(* Logix 5000 project; controller NWGG 1756-L72 rev 35.12; software revision 35.00; part 3 of 19 *)
(* tags used below, declared in another part *)
   _6Y : ALIAS FOR I25[2].3;
   _700_TREAT : ALIAS FOR I7.3;
   _709G_TREAT : ALIAS FOR B21[9].7;
   _9_DRIP_GAT : ALIAS FOR O24[7].7;
   _9_GATE_SV : ALIAS FOR O24[7].0;
   _9_GATE_SV1 : ALIAS FOR O24[7].1;
   _9_TREATER : ALIAS FOR I24[6].7;
   _9_TRT_MB : ALIAS FOR B3[9].0;
   _9_TRT_MOV : ALIAS FOR O24[7].4;
   _9_TRT_STB : ALIAS FOR B3[9].1;
   _9_TRT_STPB : ALIAS FOR B3[9].2;
   A16 : INT[250];
   A_ACC : ALIAS FOR N10[11];
   A_HOLD_B : ALIAS FOR B3[1].4;
   A_HOLD_MB : ALIAS FOR B3[1].3;
   A_HOLD_REL : ALIAS FOR B3[1].5;
   A_MAIN_CNT : ALIAS FOR C5[0].PRE;
   A_MAIN_CNT1 : ALIAS FOR C5[0].ACC;
   A_MAIN_TRE : ALIAS FOR C5[0];
   A_PRESET : ALIAS FOR N10[10];
   A_PRESET_S : ALIAS FOR N10[12];
   A_RESET_PB : ALIAS FOR B3[1].2;
   A_SET : ALIAS FOR B3[1].6;
   A_STB_AUTO : ALIAS FOR B3[1].0;
   A_STPB_AUT : ALIAS FOR B3[1].1;
   A_TREATER : ALIAS FOR I24[6].8;
   A_TREATER1 : ALIAS FOR T4[59];
   B15 : DINT[100];
   B17 : DINT[30];
   B21 : DINT[255];
   B3 : DINT[250];
   B9 : DINT[150];
   Beta : BOOL;
   C5 : COUNTER[50];
   F8 : REAL[27];
   I1 : ALIAS FOR R1S0_AENTR:1:I.Data;
   I1_000_Bit00 : ALIAS FOR I1.0;
   I1_000_Bit02 : ALIAS FOR I1.2;
   I1_000_Bit03 : ALIAS FOR I1.3;
   I1_000_Bit05 : ALIAS FOR I1.5;
   I1_000_Bit06 : ALIAS FOR I1.6;
   I1_000_Bit08 : ALIAS FOR I1.8;
   I1_000_Bit09 : ALIAS FOR I1.9;
   I1_000_Bit11 : ALIAS FOR I1.11;
   I1_000_Bit12 : ALIAS FOR I1.12;
   I1_000_Bit14 : ALIAS FOR I1.14;
   I2 : ALIAS FOR R1S0_AENTR:2:I.Data;
   I24_004_Bit00 : ALIAS FOR I24[4].0;
   I24_004_Bit01 : ALIAS FOR I24[4].1;
   I24_004_Bit02 : ALIAS FOR I24[4].2;
   I24_004_Bit03 : ALIAS FOR I24[4].3;
   I24_006_Bit13 : ALIAS FOR I24[6].13;
   I25_002_Bit04 : ALIAS FOR I25[2].4;
   I2_000_Bit00 : ALIAS FOR I2.0;
   I2_000_Bit02 : ALIAS FOR I2.2;
   I2_000_Bit03 : ALIAS FOR I2.3;
   I2_000_Bit05 : ALIAS FOR I2.5;
   I2_000_Bit06 : ALIAS FOR I2.6;
   I2_000_Bit08 : ALIAS FOR I2.8;
   I2_000_Bit09 : ALIAS FOR I2.9;
   I2_000_Bit11 : ALIAS FOR I2.11;
   I2_000_Bit12 : ALIAS FOR I2.12;
   I2_000_Bit14 : ALIAS FOR I2.14;
   I3 : ALIAS FOR R1S0_AENTR:3:I.Data;
   I3_000_Bit00 : ALIAS FOR I3.0;
   I3_000_Bit02 : ALIAS FOR I3.2;
   I3_000_Bit03 : ALIAS FOR I3.3;
   I3_000_Bit05 : ALIAS FOR I3.5;
   I3_000_Bit06 : ALIAS FOR I3.6;
   I3_000_Bit08 : ALIAS FOR I3.8;
   I3_000_Bit09 : ALIAS FOR I3.9;
   I3_000_Bit11 : ALIAS FOR I3.11;
   I3_000_Bit12 : ALIAS FOR I3.12;
   I3_000_Bit14 : ALIAS FOR I3.14;
   I4 : ALIAS FOR R1S0_AENTR:4:I.Data;
   I4_000_Bit00 : ALIAS FOR I4.0;
   I4_000_Bit02 : ALIAS FOR I4.2;
   I4_000_Bit04 : ALIAS FOR I4.4;
   InEUMax : REAL;
   MAIN_TIMER : ALIAS FOR T11[0];
   MAIN_TIMER1 : ALIAS FOR T11[1];
   N20 : DINT[30];
   N23 : DINT[5];
   N7 : DINT[100];
   O10 : ALIAS FOR R1S0_AENTR:10:O.Data;
   O11 : ALIAS FOR R1S0_AENTR:11:O.Data;
   O12 : ALIAS FOR R1S0_AENTR:12:O.Data;
   O24_005_Bit00 : ALIAS FOR O24[5].0;
   O24_005_Bit01 : ALIAS FOR O24[5].1;
   O24_005_Bit02 : ALIAS FOR O24[5].2;
   O24_007_Bit05 : ALIAS FOR O24[7].5;
   O25_010_Bit04 : ALIAS FOR O25[10].4;
   O25_010_Bit07 : ALIAS FOR O25[10].7;
   P1_AUTO_SE : ALIAS FOR B3[5].1;
   P1_RUN_AUT1 : ALIAS FOR B3[4].1;
   P1_SEC_SEL : ALIAS FOR B17[1].1;
   P2_AUTO_SE : ALIAS FOR B3[5].2;
   P2_RUN_AUT1 : ALIAS FOR B3[4].2;
   P2_SEC_SEL : ALIAS FOR B17[1].2;
   P3_AUTO_SE : ALIAS FOR B3[5].3;
   P3_RUN_AUT1 : ALIAS FOR B3[4].3;
   P3_SEC_SEL : ALIAS FOR B17[1].3;
   P4_AUTO_SE : ALIAS FOR B3[5].4;
   P4_RUN_AUT1 : ALIAS FOR B3[4].4;
   P4_SEC_SEL : ALIAS FOR B17[1].4;
   P_RESET_AU : ALIAS FOR B3[4].0;
   PUMP_NO_FL : ALIAS FOR B12[11].0;
   T11_AIRSG1 : ALIAS FOR T4[0];
   T11_AIRSG2 : ALIAS FOR T4[1];
   T11_AUTO_A : ALIAS FOR T4[61];
   T11_TREAT : ALIAS FOR B3[11].0;
   T11_TRT_MO : ALIAS FOR T4[41];
   T12_DLY_TR : ALIAS FOR T4[2];
   T12_DLY_TR3 : ALIAS FOR T4[3];
   T12_TREAT : ALIAS FOR B3[12].0;
   T12_TRT_MO : ALIAS FOR T4[42];
   T13_DLY_TR : ALIAS FOR T4[4];
   T13_DLY_TR3 : ALIAS FOR T4[5];
   T13_TREAT : ALIAS FOR B3[13].0;
   T13_TRT_MO : ALIAS FOR T4[43];
   T13C_TREAT : ALIAS FOR B21[70].10;
   T14_DLY_TR : ALIAS FOR T4[6];
   T14_DLY_TR3 : ALIAS FOR T4[7];
   T14_TREAT : ALIAS FOR B3[14].0;
   T14_TRT_MO : ALIAS FOR T4[44];
   T15_TREAT : ALIAS FOR B3[15].0;
   T15_TRT_MO : ALIAS FOR T4[45];
   T15_TRT_OF : ALIAS FOR T4[9];
   T15_TRT_ON : ALIAS FOR T4[8];
   T16_TREAT : ALIAS FOR B3[16].0;
   T16_TRT_MO : ALIAS FOR T4[46];
   T16_TRT_OF : ALIAS FOR T4[11];
   T16_TRT_ON : ALIAS FOR T4[10];

   T17_HOLD_A : ALIAS FOR B3[17].3;
   T17_HOLD_M : ALIAS FOR B3[17].6;
   T17_K_FACT : ALIAS FOR F8[13];
   T17_LOW_BI : ALIAS FOR B15[17].2;
   T17_METER : ALIAS FOR I2.5;
   T17_NO_PAS : ALIAS FOR B17[17].2;
   T17_NULL_V : ALIAS FOR A16[178];
   T17_NULL_V1 : ALIAS FOR A16[179];
   T17_OP_DEF : ALIAS FOR A16[176];
   T17_OP_DEF1 : ALIAS FOR A16[177];
   T17_OP_NAM : ALIAS FOR A16[173];
   T17_OP_NAM1 : ALIAS FOR A16[174];
   T17_OPEN_A : ALIAS FOR B3[17].8;
   T17_OPEN_M : ALIAS FOR O10.5;
   T17_OPEN_M1 : ALIAS FOR B3[17].10;
   T17_RELEAS : ALIAS FOR B3[17].5;
   T17_RESET : ALIAS FOR B3[17].7;
   T17_SET_AU : ALIAS FOR B3[17].2;
   T17_SET_DE : ALIAS FOR B3[2].6;
   T17_SET_LO : ALIAS FOR B3[17].13;
   T17_SET_MA : ALIAS FOR B3[17].12;
   T17_SET_NA : ALIAS FOR A16[170];
   T17_SET_NA1 : ALIAS FOR A16[171];
   T17_SET_NA2 : ALIAS FOR B17[17].0;
   T17_STOP_A : ALIAS FOR B3[17].4;
   T17_TREAT : ALIAS FOR B3[17].0;
   T17_TRT_MO : ALIAS FOR T4[47];
   T17_TRT_MO1 : ALIAS FOR T4[47].PRE;
   T17_TRT_MO2 : ALIAS FOR T4[47].ACC;
   T17_TRT_OF : ALIAS FOR T4[13];
   T17_TRT_OF1 : ALIAS FOR T4[13].PRE;
   T17_TRT_OF2 : ALIAS FOR T4[13].ACC;
   T17_TRT_ON : ALIAS FOR T4[12];
   T17_TRT_ON1 : ALIAS FOR T4[12].PRE;
   T17_TRT_ON2 : ALIAS FOR T4[12].ACC;
   T19 : TIMER[2] := ([0].PRE := 11000, [0].ACC := 11000, [1].PRE := 60000, [1].ACC := 60000);
   T19C_AIR_G : ALIAS FOR O12.13;
   T19C_AIR_S : ALIAS FOR B21[71].11;
   T19C_CLOSE : ALIAS FOR O12.12;
   T19C_CLOSE1 : ALIAS FOR T22[3];
   T19C_CLOSE2 : ALIAS FOR T22[3].PRE;
   T19C_CLOSE3 : ALIAS FOR T22[3].ACC;
   T19C_GATE : ALIAS FOR B21[71].0;
   T19C_GATE1 : ALIAS FOR B21[71].1;
   T19C_GATE2 : ALIAS FOR B21[71].3;
   T19C_GATE3 : ALIAS FOR B21[71].4;
   T19C_GATE4 : ALIAS FOR B21[71].5;
   T19C_GATE5 : ALIAS FOR B21[71].6;
   T19C_GATE6 : ALIAS FOR B21[71].7;
   T19C_GATE7 : ALIAS FOR B21[71].8;
   T19C_GATE8 : ALIAS FOR B21[71].9;
   T19C_GATEC : ALIAS FOR B21[71].2;
   T19C_GATET : ALIAS FOR C5[4];
   T19C_OPEN : ALIAS FOR O12.11;
   T19C_SET_D : ALIAS FOR B21[71].14;
   T19C_TMR_A : ALIAS FOR C5[4].ACC;
   T19C_TMR_P : ALIAS FOR C5[4].PRE;
   T19C_TREAT : ALIAS FOR B21[71].10;
   T19C_TRT_M : ALIAS FOR T22[4];
   T19C_TRT_M1 : ALIAS FOR T22[4].PRE;
   T19C_TRT_M2 : ALIAS FOR T22[4].ACC;
   T19C_TRT_O : ALIAS FOR T22[0];
   T19C_TRT_O1 : ALIAS FOR T22[0].PRE;
   T19C_TRT_O2 : ALIAS FOR T22[0].ACC;
   T21_AIR_GA : ALIAS FOR I2.6;
   T21_AIR_SV : ALIAS FOR O10.6;
   T21_ASCII : ALIAS FOR B17[21].1;
   T21_ASSII : ALIAS FOR A16[212];
   T21_ASSII1 : ALIAS FOR A16[215];
   T21_AUTO_A : ALIAS FOR T4[71];
   T21_AUTO_A1 : ALIAS FOR T4[71].PRE;
   T21_AUTO_A2 : ALIAS FOR T4[71].ACC;
   T21_AUTO_M : ALIAS FOR B3[21].1;
   T21_AUTO_S : ALIAS FOR B3[21].14;
   T21_BINDIC : ALIAS FOR I1.1;
   T21_CAL_CL : ALIAS FOR B15[61].3;
   T21_CAL_LA : ALIAS FOR B15[61].2;
   T21_CAL_OP : ALIAS FOR B15[61].4;
   T21_CAL_ST : ALIAS FOR B15[61].1;
   T21_CLOSE : ALIAS FOR O10.7;
   T21_CLOSE1 : ALIAS FOR B3[21].9;
   T21_CLOSE2 : ALIAS FOR B3[21].11;
   T21_CORREC : ALIAS FOR F8[16];
   T21_FAULT : ALIAS FOR B3[21].15;
   T21_GATE_C : ALIAS FOR C5[21];
   T21_GATE_C1 : ALIAS FOR C5[21].PRE;
   T21_GATE_C2 : ALIAS FOR C5[21].ACC;
   T21_HOLD_A : ALIAS FOR B3[21].3;
   T21_HOLD_M : ALIAS FOR B3[21].6;
   T21_K_FACT : ALIAS FOR F8[15];
   T21_LOW_BI : ALIAS FOR B15[21].2;
   T21_METER : ALIAS FOR I2.8;
   T21_MOVE_D : ALIAS FOR I2.7;
   T21_NO_PAS : ALIAS FOR B17[21].2;
   T21_NULL_V : ALIAS FOR A16[218];
   T21_NULL_V1 : ALIAS FOR A16[219];
   T21_OP_DEF : ALIAS FOR A16[216];
   T21_OP_DEF1 : ALIAS FOR A16[217];
   T21_OP_NAM : ALIAS FOR A16[213];
   T21_OP_NAM1 : ALIAS FOR A16[214];
   T21_OPEN_A : ALIAS FOR B3[21].8;
   T21_OPEN_M : ALIAS FOR O10.8;
   T21_OPEN_M1 : ALIAS FOR B3[21].10;
   T21_RELEAS : ALIAS FOR B3[21].5;
   T21_RESET : ALIAS FOR B3[21].7;
   T21_SET_AU : ALIAS FOR B3[21].2;
   T21_SET_DE : ALIAS FOR B3[2].7;
   T21_SET_LO : ALIAS FOR B3[21].13;
   T21_SET_MA : ALIAS FOR B3[21].12;
   T21_SET_NA : ALIAS FOR A16[210];
   T21_SET_NA1 : ALIAS FOR A16[211];
   T21_SET_NA2 : ALIAS FOR B17[21].0;
   T21_STOP_A : ALIAS FOR B3[21].4;
   T21_TREAT : ALIAS FOR B3[21].0;
   T21_TRT_MO : ALIAS FOR T4[48];
   T21_TRT_MO1 : ALIAS FOR T4[48].PRE;
   T21_TRT_MO2 : ALIAS FOR T4[48].ACC;
   T21_TRT_OF : ALIAS FOR T4[15];
   T21_TRT_OF1 : ALIAS FOR T4[15].PRE;
   T21_TRT_OF2 : ALIAS FOR T4[15].ACC;
   T21_TRT_ON : ALIAS FOR T4[14];
   T21_TRT_ON1 : ALIAS FOR T4[14].PRE;
   T21_TRT_ON2 : ALIAS FOR T4[14].ACC;
   T22 : TIMER[100] := ([0].PRE := 1000, [1].PRE := 10000, [1].ACC := 10000, [2].PRE := 10000, [2].ACC := 10000, [3].PRE := 1000, [3].ACC := 1000, [4].PRE := 2500, [5].PRE := 7000, [6].PRE := 10000, [6].ACC := 10000, [7].PRE := 2500, [8].PRE := 1000, [8].ACC := 1000, [9].PRE := 1000, [9].ACC := 1000, [10].PRE := 2000, [13].PRE := 10000, [14].PRE := 10000, [15].PRE := 10000, [16].PRE := 10000, [17].PRE := 10000);
   T22_AIR_GA : ALIAS FOR I2.9;
   T22_AIR_SV : ALIAS FOR O10.9;
   T22_ASCII : ALIAS FOR B17[22].1;
   T22_ASSII : ALIAS FOR A16[222];
   T22_ASSII1 : ALIAS FOR A16[225];
   T22_AUTO_A : ALIAS FOR T4[72];
   T22_AUTO_A1 : ALIAS FOR T4[72].PRE;
   T22_AUTO_A2 : ALIAS FOR T4[72].ACC;
   T22_AUTO_M : ALIAS FOR B3[22].1;
   T22_AUTO_S : ALIAS FOR B3[22].14;
   T22_BINDIC : ALIAS FOR I1.4;
   T22_CAL_CL : ALIAS FOR B15[62].3;
   T22_CAL_LA : ALIAS FOR B15[62].2;
   T22_CAL_OP : ALIAS FOR B15[62].4;
   T22_CAL_ST : ALIAS FOR B15[62].1;
   T22_CLOSE : ALIAS FOR O10.10;
   T22_CLOSE1 : ALIAS FOR B3[22].9;
   T22_CLOSE2 : ALIAS FOR B3[22].11;
   T22_CORREC : ALIAS FOR F8[18];
   T22_FAULT : ALIAS FOR B3[22].15;
   T22_GATE_C : ALIAS FOR C5[22];
   T22_GATE_C1 : ALIAS FOR C5[22].PRE;
   T22_GATE_C2 : ALIAS FOR C5[22].ACC;
   T22_HOLD_A : ALIAS FOR B3[22].3;
   T22_HOLD_M : ALIAS FOR B3[22].6;
   T22_K_FACT : ALIAS FOR F8[17];
   T22_LOW_BI : ALIAS FOR B15[22].2;
   T22_METER : ALIAS FOR I2.11;
   T22_MOVE_D : ALIAS FOR I2.10;
   T22_NO_PAS : ALIAS FOR B17[22].2;
   T22_NULL_V : ALIAS FOR A16[228];
   T22_NULL_V1 : ALIAS FOR A16[229];
   T22_OP_DEF : ALIAS FOR A16[226];
   T22_OP_DEF1 : ALIAS FOR A16[227];
   T22_OP_NAM : ALIAS FOR A16[223];
   T22_OP_NAM1 : ALIAS FOR A16[224];
   T22_OPEN_A : ALIAS FOR B3[22].8;
   T22_OPEN_M : ALIAS FOR O10.11;
   T22_OPEN_M1 : ALIAS FOR B3[22].10;
   T22_RELEAS : ALIAS FOR B3[22].5;
   T22_RESET : ALIAS FOR B3[22].7;
   T22_SET_AU : ALIAS FOR B3[22].2;
   T22_SET_DE : ALIAS FOR B3[2].8;
   T22_SET_LO : ALIAS FOR B3[22].13;
   T22_SET_MA : ALIAS FOR B3[22].12;
   T22_SET_NA : ALIAS FOR A16[220];
   T22_SET_NA1 : ALIAS FOR A16[221];
   T22_SET_NA2 : ALIAS FOR B17[22].0;
   T22_STOP_A : ALIAS FOR B3[22].4;
   T22_TREAT : ALIAS FOR B3[22].0;
   T22_TRT_MO : ALIAS FOR T4[49];
   T22_TRT_MO1 : ALIAS FOR T4[49].PRE;
   T22_TRT_MO2 : ALIAS FOR T4[49].ACC;
   T22_TRT_OF : ALIAS FOR T4[17];
   T22_TRT_OF1 : ALIAS FOR T4[17].PRE;
   T22_TRT_OF2 : ALIAS FOR T4[17].ACC;
   T22_TRT_ON : ALIAS FOR T4[16];
   T22_TRT_ON1 : ALIAS FOR T4[16].PRE;
   T22_TRT_ON2 : ALIAS FOR T4[16].ACC;
   T23_AIR_GA : ALIAS FOR I2.12;
   T23_AIR_SV : ALIAS FOR O10.12;
   T23_ASCII : ALIAS FOR B17[23].1;
   T23_ASSII : ALIAS FOR A16[232];
   T23_ASSII1 : ALIAS FOR A16[235];
   T23_AUTO_A : ALIAS FOR T4[73];
   T23_AUTO_A1 : ALIAS FOR T4[73].PRE;
   T23_AUTO_A2 : ALIAS FOR T4[73].ACC;
   T23_AUTO_M : ALIAS FOR B3[23].1;
   T23_AUTO_S : ALIAS FOR B3[23].14;
   T23_BINDIC : ALIAS FOR I1.7;
   T23_CAL_CL : ALIAS FOR B15[63].3;
   T23_CAL_LA : ALIAS FOR B15[63].2;
   T23_CAL_OP : ALIAS FOR B15[63].4;
   T23_CAL_ST : ALIAS FOR B15[63].1;
   T23_CLOSE : ALIAS FOR O10.13;
   T23_CLOSE1 : ALIAS FOR B3[23].9;
   T23_CLOSE2 : ALIAS FOR B3[23].11;
   T23_CORREC : ALIAS FOR F8[20];
   T23_FAULT : ALIAS FOR B3[23].15;
   T23_GATE_C : ALIAS FOR C5[23];
   T23_GATE_C1 : ALIAS FOR C5[23].PRE;
   T23_GATE_C2 : ALIAS FOR C5[23].ACC;
   T23_HOLD_A : ALIAS FOR B3[23].3;
   T23_HOLD_M : ALIAS FOR B3[23].6;
   T23_K_FACT : ALIAS FOR F8[19];
   T23_LOW_BI : ALIAS FOR B15[23].2;
   T23_METER : ALIAS FOR I2.14;
   T23_MOVE_D : ALIAS FOR I2.13;
   T23_NO_PAS : ALIAS FOR B17[23].2;
   T23_NULL_V : ALIAS FOR A16[238];
   T23_NULL_V1 : ALIAS FOR A16[239];
   T23_OP_DEF : ALIAS FOR A16[236];
   T23_OP_DEF1 : ALIAS FOR A16[237];
   T23_OP_NAM : ALIAS FOR A16[233];
   T23_OP_NAM1 : ALIAS FOR A16[234];
   T23_OPEN_A : ALIAS FOR B3[23].8;
   T23_OPEN_M : ALIAS FOR O10.14;
   T23_OPEN_M1 : ALIAS FOR B3[23].10;
   T23_RELEAS : ALIAS FOR B3[23].5;
   T23_RESET : ALIAS FOR B3[23].7;
   T23_SET_AU : ALIAS FOR B3[23].2;
   T23_SET_DE : ALIAS FOR B3[2].9;
   T23_SET_LO : ALIAS FOR B3[23].13;
   T23_SET_MA : ALIAS FOR B3[23].12;
   T23_SET_NA : ALIAS FOR A16[230];
   T23_SET_NA1 : ALIAS FOR A16[231];
   T23_SET_NA2 : ALIAS FOR B17[23].0;
   T23_STOP_A : ALIAS FOR B3[23].4;
   T23_TREAT : ALIAS FOR B3[23].0;
   T23_TRT_MO : ALIAS FOR T4[50];
   T23_TRT_MO1 : ALIAS FOR T4[50].PRE;
   T23_TRT_MO2 : ALIAS FOR T4[50].ACC;
   T23_TRT_OF : ALIAS FOR T4[19];
   T23_TRT_OF1 : ALIAS FOR T4[19].PRE;
   T23_TRT_OF2 : ALIAS FOR T4[19].ACC;
   T23_TRT_ON : ALIAS FOR T4[18];
   T23_TRT_ON1 : ALIAS FOR T4[18].PRE;
   T23_TRT_ON2 : ALIAS FOR T4[18].ACC;
   T24_AIR_GA : ALIAS FOR I3.0;
   T24_AIR_SV : ALIAS FOR O11.0;
   T24_ASCII : ALIAS FOR B17[24].1;
   T24_ASSII : ALIAS FOR A16[242];
   T24_ASSII1 : ALIAS FOR A16[245];
   T24_AUTO_A : ALIAS FOR T4[74];
   T24_AUTO_A1 : ALIAS FOR T4[74].PRE;
   T24_AUTO_A2 : ALIAS FOR T4[74].ACC;
   T24_AUTO_M : ALIAS FOR B3[24].1;
   T24_AUTO_S : ALIAS FOR B3[24].14;
   T24_BINDIC : ALIAS FOR I1.10;
   T24_CAL_CL : ALIAS FOR B15[64].3;
   T24_CAL_LA : ALIAS FOR B15[64].2;
   T24_CAL_OP : ALIAS FOR B15[64].4;
   T24_CAL_ST : ALIAS FOR B15[64].1;
   T24_CLOSE : ALIAS FOR O11.1;
   T24_CLOSE1 : ALIAS FOR B3[24].9;
   T24_CLOSE2 : ALIAS FOR B3[24].11;
   T24_CORREC : ALIAS FOR F8[22];
   T24_FAULT : ALIAS FOR B3[24].15;
   T24_GATE_C : ALIAS FOR C5[24];
   T24_GATE_C1 : ALIAS FOR C5[24].PRE;
   T24_GATE_C2 : ALIAS FOR C5[24].ACC;
   T24_HOLD_A : ALIAS FOR B3[24].3;
   T24_HOLD_M : ALIAS FOR B3[24].6;
   T24_K_FACT : ALIAS FOR F8[21];
   T24_LOW_BI : ALIAS FOR B15[24].2;
   T24_METER : ALIAS FOR I3.2;
   T24_MOVE_D : ALIAS FOR I3.1;
   T24_NO_PAS : ALIAS FOR B17[24].2;
   T24_NULL_V : ALIAS FOR A16[248];
   T24_NULL_V1 : ALIAS FOR A16[249];
   T24_OP_DEF : ALIAS FOR A16[246];
   T24_OP_DEF1 : ALIAS FOR A16[247];
   T24_OP_NAM : ALIAS FOR A16[243];
   T24_OP_NAM1 : ALIAS FOR A16[244];
   T24_OPEN_A : ALIAS FOR B3[24].8;
   T24_OPEN_M : ALIAS FOR O11.2;
   T24_OPEN_M1 : ALIAS FOR B3[24].10;
   T24_RELEAS : ALIAS FOR B3[24].5;
   T24_RESET : ALIAS FOR B3[24].7;
   T24_SET_AU : ALIAS FOR B3[24].2;
   T24_SET_DE : ALIAS FOR B3[2].10;
   T24_SET_LO : ALIAS FOR B3[24].13;
   T24_SET_MA : ALIAS FOR B3[24].12;
   T24_SET_NA : ALIAS FOR A16[240];
   T24_SET_NA1 : ALIAS FOR A16[241];
   T24_SET_NA2 : ALIAS FOR B17[24].0;
   T24_STOP_A : ALIAS FOR B3[24].4;
   T24_TREAT : ALIAS FOR B3[24].0;
   T24_TRT_MO : ALIAS FOR T4[51];
   T24_TRT_MO1 : ALIAS FOR T4[51].PRE;
   T24_TRT_MO2 : ALIAS FOR T4[51].ACC;
   T24_TRT_OF : ALIAS FOR T4[21];
   T24_TRT_OF1 : ALIAS FOR T4[21].PRE;
   T24_TRT_OF2 : ALIAS FOR T4[21].ACC;
   T24_TRT_ON : ALIAS FOR T4[20];
   T24_TRT_ON1 : ALIAS FOR T4[20].PRE;
   T24_TRT_ON2 : ALIAS FOR T4[20].ACC;
   T25 : TIMER[9] := ([0].PRE := 1000, [0].ACC := 1000, [1].PRE := 10, [1].ACC := 10, [2].PRE := 1000, [2].ACC := 1000, [3].PRE := 10, [3].ACC := 10, [4].PRE := 5000, [4].ACC := 5000, [5].PRE := 5000, [5].ACC := 5000, [6].PRE := 60000, [6].ACC := 60000, [7].PRE := 1000, [7].ACC := 1000);
   T25_AIR_GA : ALIAS FOR I3.3;
   T25_AIR_SV : ALIAS FOR O11.3;
   T25_ASCII : ALIAS FOR B17[25].1;
   T25_ASSII : ALIAS FOR A16[192];
   T25_ASSII1 : ALIAS FOR A16[195];
   T25_AUTO_A : ALIAS FOR T4[75];
   T25_AUTO_A1 : ALIAS FOR T4[75].PRE;
   T25_AUTO_A2 : ALIAS FOR T4[75].ACC;
   T25_AUTO_M : ALIAS FOR B3[25].1;
   T25_AUTO_S : ALIAS FOR B3[25].14;
   T25_BINDIC : ALIAS FOR I1.13;
   T25_CAL_CL : ALIAS FOR B15[65].3;
   T25_CAL_LA : ALIAS FOR B15[65].2;
   T25_CAL_OP : ALIAS FOR B15[65].4;
   T25_CAL_ST : ALIAS FOR B15[65].1;
   T25_CLOSE : ALIAS FOR O11.4;
   T25_CLOSE1 : ALIAS FOR B3[25].9;
   T25_CLOSE2 : ALIAS FOR B3[25].11;
   T25_CORREC : ALIAS FOR F8[24];
   T25_FAULT : ALIAS FOR B3[25].15;
   T25_GATE_C : ALIAS FOR C5[25];
   T25_GATE_C1 : ALIAS FOR C5[25].PRE;
   T25_GATE_C2 : ALIAS FOR C5[25].ACC;
   T25_HOLD_A : ALIAS FOR B3[25].3;
   T25_HOLD_M : ALIAS FOR B3[25].6;
   T25_K_FACT : ALIAS FOR F8[23];
   T25_LOW_BI : ALIAS FOR B15[25].2;
   T25_METER : ALIAS FOR I3.5;
   T25_MOVE_D : ALIAS FOR I3.4;
   T25_NO_PAS : ALIAS FOR B17[25].2;
   T25_NULL_V : ALIAS FOR A16[198];
   T25_NULL_V1 : ALIAS FOR A16[199];
   T25_OP_DEF : ALIAS FOR A16[196];
   T25_OP_DEF1 : ALIAS FOR A16[197];
   T25_OP_NAM : ALIAS FOR A16[193];
   T25_OP_NAM1 : ALIAS FOR A16[194];
   T25_OPEN_A : ALIAS FOR B3[25].8;
   T25_OPEN_M : ALIAS FOR O11.5;
   T25_OPEN_M1 : ALIAS FOR B3[25].10;
   T25_RELEAS : ALIAS FOR B3[25].5;
   T25_RESET : ALIAS FOR B3[25].7;
   T25_SET_AU : ALIAS FOR B3[25].2;
   T25_SET_DE : ALIAS FOR B3[2].11;
   T25_SET_LO : ALIAS FOR B3[25].13;
   T25_SET_MA : ALIAS FOR B3[25].12;
   T25_SET_NA : ALIAS FOR A16[190];
   T25_SET_NA1 : ALIAS FOR A16[191];
   T25_SET_NA2 : ALIAS FOR B17[25].0;
   T25_STOP_A : ALIAS FOR B3[25].4;
   T25_TREAT : ALIAS FOR B3[25].0;
   T25_TRT_MO : ALIAS FOR T4[52];
   T25_TRT_MO1 : ALIAS FOR T4[52].PRE;
   T25_TRT_MO2 : ALIAS FOR T4[52].ACC;
   T25_TRT_OF : ALIAS FOR T4[23];
   T25_TRT_OF1 : ALIAS FOR T4[23].PRE;
   T25_TRT_OF2 : ALIAS FOR T4[23].ACC;
   T25_TRT_ON : ALIAS FOR T4[22];
   T25_TRT_ON1 : ALIAS FOR T4[22].PRE;
   T25_TRT_ON2 : ALIAS FOR T4[22].ACC;
   T26_AIR_GA : ALIAS FOR I3.6;
   T26_AIR_SV : ALIAS FOR O11.6;
   T26_ASCII : ALIAS FOR B17[26].1;
   T26_ASSII : ALIAS FOR A16[202];
   T26_ASSII1 : ALIAS FOR A16[205];
   T26_AUTO_A : ALIAS FOR T4[76];
   T26_AUTO_A1 : ALIAS FOR T4[76].PRE;
   T26_AUTO_A2 : ALIAS FOR T4[76].ACC;
   T26_AUTO_M : ALIAS FOR B3[26].1;
   T26_AUTO_S : ALIAS FOR B3[26].14;
   T26_BINDIC : ALIAS FOR I1.15;
   T26_CAL_CL : ALIAS FOR B15[66].3;
   T26_CAL_LA : ALIAS FOR B15[66].2;
   T26_CAL_OP : ALIAS FOR B15[66].4;
   T26_CAL_ST : ALIAS FOR B15[66].1;
   T26_CLOSE : ALIAS FOR O11.7;
   T26_CLOSE1 : ALIAS FOR B3[26].9;
   T26_CLOSE2 : ALIAS FOR B3[26].11;
   T26_CORREC : ALIAS FOR F8[26];
   T26_FAULT : ALIAS FOR B3[26].15;
   T26_GATE_C : ALIAS FOR C5[26];
   T26_GATE_C1 : ALIAS FOR C5[26].PRE;
   T26_GATE_C2 : ALIAS FOR C5[26].ACC;
   T26_HOLD_A : ALIAS FOR B3[26].3;
   T26_HOLD_M : ALIAS FOR B3[26].6;
   T26_K_FACT : ALIAS FOR F8[25];
   T26_LOW_BI : ALIAS FOR B15[26].2;
   T26_METER : ALIAS FOR I3.8;
   T26_MOVE_D : ALIAS FOR I3.7;
   T26_NO_PAS : ALIAS FOR B17[26].2;
   T26_NULL_V : ALIAS FOR A16[208];
   T26_NULL_V1 : ALIAS FOR A16[209];
   T26_OP_DEF : ALIAS FOR A16[206];
   T26_OP_DEF1 : ALIAS FOR A16[207];
   T26_OP_NAM : ALIAS FOR A16[203];
   T26_OP_NAM1 : ALIAS FOR A16[204];
   T26_OPEN_A : ALIAS FOR B3[26].8;
   T26_OPEN_M : ALIAS FOR O11.8;
   T26_OPEN_M1 : ALIAS FOR B3[26].10;
   T26_RELEAS : ALIAS FOR B3[26].5;
   T26_RESET : ALIAS FOR B3[26].7;
   T26_SET_AU : ALIAS FOR B3[26].2;
   T26_SET_DE : ALIAS FOR B3[2].12;
   T26_SET_LO : ALIAS FOR B3[26].13;
   T26_SET_MA : ALIAS FOR B3[26].12;
   T26_SET_NA : ALIAS FOR A16[200];
   T26_SET_NA1 : ALIAS FOR A16[201];
   T26_SET_NA2 : ALIAS FOR B17[26].0;
   T26_STOP_A : ALIAS FOR B3[26].4;
   T26_TREAT : ALIAS FOR B3[26].0;
   T26_TRT_MO : ALIAS FOR T4[53];
   T26_TRT_MO1 : ALIAS FOR T4[53].PRE;
   T26_TRT_MO2 : ALIAS FOR T4[53].ACC;
   T26_TRT_OF : ALIAS FOR T4[25];
   T26_TRT_OF1 : ALIAS FOR T4[25].PRE;
   T26_TRT_OF2 : ALIAS FOR T4[25].ACC;
   T26_TRT_ON : ALIAS FOR T4[24];
   T26_TRT_ON1 : ALIAS FOR T4[24].PRE;
   T26_TRT_ON2 : ALIAS FOR T4[24].ACC;
   T27_AIR_GA : ALIAS FOR I3.9;
   T27_AIR_SV : ALIAS FOR O11.9;
   T27_AUTO_A : ALIAS FOR T4[77];
   T27_AUTO_A1 : ALIAS FOR T4[77].PRE;
   T27_AUTO_A2 : ALIAS FOR T4[77].ACC;
   T27_AUTO_M : ALIAS FOR B3[27].1;
   T27_AUTO_S : ALIAS FOR B3[27].14;
   T27_CLOSE : ALIAS FOR O11.10;
   T27_CLOSE1 : ALIAS FOR B3[27].9;
   T27_CLOSE2 : ALIAS FOR B3[27].11;
   T27_FAULT : ALIAS FOR B3[27].15;
   T27_GATE_C : ALIAS FOR C5[27];
   T27_GATE_C1 : ALIAS FOR C5[27].PRE;
   T27_GATE_C2 : ALIAS FOR C5[27].ACC;
   T27_HOLD_A : ALIAS FOR B3[27].3;
   T27_HOLD_M : ALIAS FOR B3[27].6;
   T27_LOW_BI : ALIAS FOR B15[27].2;
   T27_METER : ALIAS FOR I3.11;
   T27_OPEN_A : ALIAS FOR B3[27].8;
   T27_OPEN_M : ALIAS FOR O11.11;
   T27_OPEN_M1 : ALIAS FOR B3[27].10;
   T27_RELEAS : ALIAS FOR B3[27].5;
   T27_RESET : ALIAS FOR B3[27].7;
   T27_SET_AU : ALIAS FOR B3[27].2;
   T27_SET_DE : ALIAS FOR B3[2].13;
   T27_SET_LO : ALIAS FOR B3[27].13;
   T27_SET_MA : ALIAS FOR B3[27].12;
   T27_STOP_A : ALIAS FOR B3[27].4;
   T27_TREAT : ALIAS FOR B3[27].0;
   T27_TRT_MO : ALIAS FOR T4[54];
   T27_TRT_MO1 : ALIAS FOR T4[54].PRE;
   T27_TRT_MO2 : ALIAS FOR T4[54].ACC;
   T27_TRT_OF : ALIAS FOR T4[27];
   T27_TRT_OF1 : ALIAS FOR T4[27].PRE;
   T27_TRT_OF2 : ALIAS FOR T4[27].ACC;
   T27_TRT_ON : ALIAS FOR T4[26];
   T27_TRT_ON1 : ALIAS FOR T4[26].PRE;
   T27_TRT_ON2 : ALIAS FOR T4[26].ACC;
   T28_AIR_SV : ALIAS FOR O11.12;
   T28_AUTO_A : ALIAS FOR T4[78];
   T28_AUTO_A1 : ALIAS FOR T4[78].PRE;
   T28_AUTO_A2 : ALIAS FOR T4[78].ACC;
   T28_AUTO_M : ALIAS FOR B3[28].1;
   T28_AUTO_S : ALIAS FOR B3[28].14;
   T28_CLOSE : ALIAS FOR O11.13;
   T28_CLOSE1 : ALIAS FOR B3[28].9;
   T28_CLOSE2 : ALIAS FOR B3[28].11;
   T28_FAULT : ALIAS FOR B3[28].15;
   T28_GATE_C : ALIAS FOR C5[28];
   T28_GATE_C1 : ALIAS FOR C5[28].PRE;
   T28_GATE_C2 : ALIAS FOR C5[28].ACC;
   T28_GATE_O : ALIAS FOR I3.12;
   T28_HOLD_A : ALIAS FOR B3[28].3;
   T28_HOLD_M : ALIAS FOR B3[28].6;
   T28_LOW_BI : ALIAS FOR B15[28].2;
   T28_METER : ALIAS FOR I3.14;
   T28_OPEN_A : ALIAS FOR B3[28].8;
   T28_OPEN_M : ALIAS FOR O11.14;
   T28_OPEN_M1 : ALIAS FOR B3[28].10;
   T28_RELEAS : ALIAS FOR B3[28].5;
   T28_RESET : ALIAS FOR B3[28].7;
   T28_SET_AU : ALIAS FOR B3[28].2;
   T28_SET_DE : ALIAS FOR B3[2].14;
   T28_SET_LO : ALIAS FOR B3[28].13;
   T28_SET_MA : ALIAS FOR B3[28].12;
   T28_STOP_A : ALIAS FOR B3[28].4;
   T28_TREAT : ALIAS FOR B3[28].0;
   T28_TRT_MO : ALIAS FOR T4[55];
   T28_TRT_MO1 : ALIAS FOR T4[55].PRE;
   T28_TRT_MO2 : ALIAS FOR T4[55].ACC;
   T28_TRT_OF : ALIAS FOR T4[29];
   T28_TRT_OF1 : ALIAS FOR T4[29].PRE;
   T28_TRT_OF2 : ALIAS FOR T4[29].ACC;
   T28_TRT_ON : ALIAS FOR T4[28];
   T28_TRT_ON1 : ALIAS FOR T4[28].PRE;
   T28_TRT_ON2 : ALIAS FOR T4[28].ACC;
   T29_AIR_GA : ALIAS FOR I4.0;
   T29_AIR_SV : ALIAS FOR O12.0;
   T29_AUTO_A : ALIAS FOR T4[79];
   T29_AUTO_A1 : ALIAS FOR T4[79].PRE;
   T29_AUTO_A2 : ALIAS FOR T4[79].ACC;
   T29_AUTO_M : ALIAS FOR B3[29].1;
   T29_AUTO_S : ALIAS FOR B3[29].14;
   T29_CLOSE : ALIAS FOR O12.1;
   T29_CLOSE1 : ALIAS FOR B3[29].9;
   T29_CLOSE2 : ALIAS FOR B3[29].11;
   T29_FAULT : ALIAS FOR B3[29].15;
   T29_GATE_C : ALIAS FOR C5[29];
   T29_GATE_C1 : ALIAS FOR C5[29].PRE;
   T29_GATE_C2 : ALIAS FOR C5[29].ACC;
   T29_HOLD_A : ALIAS FOR B3[29].3;
   T29_HOLD_M : ALIAS FOR B3[29].6;
   T29_LOW_BI : ALIAS FOR B15[29].2;
   T29_METER : ALIAS FOR I4.2;
   T29_OPEN_A : ALIAS FOR B3[29].8;
   T29_OPEN_M : ALIAS FOR O12.2;
   T29_OPEN_M1 : ALIAS FOR B3[29].10;
   T29_RELEAS : ALIAS FOR B3[29].5;
   T29_RESET : ALIAS FOR B3[29].7;
   T29_SET_AU : ALIAS FOR B3[29].2;
   T29_SET_DE : ALIAS FOR B3[2].15;
   T29_SET_LO : ALIAS FOR B3[29].13;
   T29_SET_MA : ALIAS FOR B3[29].12;
   T29_STOP_A : ALIAS FOR B3[29].4;
   T29_TREAT : ALIAS FOR B3[29].0;
   T29_TRT_MO : ALIAS FOR T4[56];
   T29_TRT_MO1 : ALIAS FOR T4[56].PRE;
   T29_TRT_MO2 : ALIAS FOR T4[56].ACC;
   T29_TRT_OF : ALIAS FOR T4[31];
   T29_TRT_OF1 : ALIAS FOR T4[31].PRE;
   T29_TRT_OF2 : ALIAS FOR T4[31].ACC;
   T29_TRT_ON : ALIAS FOR T4[30];
   T29_TRT_ON1 : ALIAS FOR T4[30].PRE;
   T29_TRT_ON2 : ALIAS FOR T4[30].ACC;
   T4 : TIMER[100] := ([0].PRE := 18000, [1].PRE := 18000, [1].ACC := 18000, [2].PRE := 11000, [3].PRE := 16000, [3].ACC := 16004, [4].PRE := 10000, [5].PRE := 16000, [5].ACC := 16000, [6].PRE := 9000, [7].PRE := 16000, [7].ACC := 16000, [8].PRE := 9000, [9].PRE := 14000, [9].ACC := 14000, [10].PRE := 11000, [11].PRE := 13000, [11].ACC := 13000, [12].PRE := 9000, [13].PRE := 13000, [13].ACC := 13000, [14].PRE := 12000, [15].PRE := 17000, [15].ACC := 17000, [16].PRE := 16000, [17].PRE := 21000, [17].ACC := 21015, [18].PRE := 20000, [19].PRE := 24000, [19].ACC := 24000, [20].PRE := 16000, [21].PRE := 21000, [21].ACC := 21000, [22].PRE := 20000, [23].PRE := 21000, [23].ACC := 21000, [24].PRE := 23000, [25].PRE := 26000, [25].ACC := 26000, [26].PRE := 26000, [27].PRE := 25000, [27].ACC := 25000, [28].PRE := 30000, [29].PRE := 29000, [29].ACC := 29000, [30].PRE := 33000, [31].PRE := 33000, [31].ACC := 33000, [32].PRE := 60000, [33].PRE := 250, [33].ACC := 251, [34].PRE := 1500000, [34].EN := 1, [34].DN := 1, [35].ACC := 2, [35].EN := 1, [35].DN := 1, [36].PRE := 3000, [36].ACC := 3001, [36].EN := 1,
        [36].DN := 1, [37].PRE := 3000, [37].ACC := 3001, [37].EN := 1, [37].DN := 1, [38].PRE := 3000, [38].ACC := 3001, [38].EN := 1, [38].DN := 1, [39].PRE := 3000, [39].ACC := 3001, [39].EN := 1, [39].DN := 1, [40].PRE := 3000, [40].ACC := 3001, [40].EN := 1, [40].DN := 1, [41].PRE := 2500, [42].PRE := 2500, [43].PRE := 2500, [44].PRE := 2500, [45].PRE := 2500, [46].PRE := 2500, [47].PRE := 2500, [48].PRE := 2500, [49].PRE := 2500, [50].PRE := 2500, [51].PRE := 2500, [52].PRE := 2500, [53].PRE := 2500, [54].PRE := 2500, [55].PRE := 2500, [56].PRE := 2500, [57].PRE := 3000, [57].ACC := 3001, [57].EN := 1, [57].DN := 1, [58].PRE := 3000, [58].ACC := 3001, [58].EN := 1, [58].DN := 1, [59].PRE := 1000, [59].ACC := 1000, [60].PRE := 1000, [61].PRE := 30000, [61].ACC := 30000, [63].PRE := 30, [64].PRE := 30, [81].PRE := 30000, [82].PRE := 30000, [83].PRE := 30000, [84].PRE := 30000, [85].PRE := 30000, [86].PRE := 30000, [87].PRE := 30000, [88].PRE := 30000, [89].PRE := 30000, [90].PRE := 30000, [91].PRE := 30000, [92].PRE := 30000,
        [93].PRE := 30000, [94].PRE := 30000, [95].PRE := 30000, [96].PRE := 30000, [97].PRE := 30000, [99].PRE := 30000);
   T41_CLOSE : ALIAS FOR O12.3;
   T41_CLOSE1 : ALIAS FOR B3[41].1;
   T41_OPEN_G : ALIAS FOR B3[41].0;
   T41_OPEN_M : ALIAS FOR O12.4;
   T41_SLIDE : ALIAS FOR I4.3;
   T42_CLOSE : ALIAS FOR O12.5;
   T42_CLOSE1 : ALIAS FOR B3[42].1;
   T42_OPEN_G : ALIAS FOR B3[42].0;
   T42_OPEN_M : ALIAS FOR O12.6;
   T42_SLIDE : ALIAS FOR I4.5;
   test : BOOL;
   testbit : BOOL := 1;
   testCounter : COUNTER;
   testint : DINT;
   TestOneshot : BOOL := 1;
   TestOneshow : BOOL;
   testOutput : BOOL;
   TestOutputBit : BOOL;
   testStorageBit : BOOL;
   TestTag : REAL;
   testTmrOffDelay : TIMER := (PRE := 5000, ACC := 5000);
   textctr : COUNTER := (DN := 1);
   TicketTreatPumpActive : DINT;
   TicketTreatPumpSet : DINT;
   TK11_COLOR : ALIAS FOR N7[50];
   TK11_PUMP : ALIAS FOR N7[70];
   TK12_COLOR : ALIAS FOR N7[51];
   TK12_PUMP : ALIAS FOR N7[71];
   TK13_COLOR : ALIAS FOR N7[52];
   TK13_PUMP : ALIAS FOR N7[72];
   TK14_COLOR : ALIAS FOR N7[53];
   TK14_PUMP : ALIAS FOR N7[73];
   TK15_COLOR : ALIAS FOR N7[54];
   TK15_PUMP : ALIAS FOR N7[74];
   TK16_COLOR : ALIAS FOR N7[55];
   TK16_PUMP : ALIAS FOR N7[75];
   TK17_COLOR : ALIAS FOR N7[56];
   TK17_PUMP : ALIAS FOR N7[76];
   TK21_COLOR : ALIAS FOR N7[57];
   TK21_PUMP : ALIAS FOR N7[77];
   TK22_COLOR : ALIAS FOR N7[58];
   TK22_PUMP : ALIAS FOR N7[78];
   TK23_COLOR : ALIAS FOR N7[59];
   TK23_PUMP : ALIAS FOR N7[79];
   TK24_COLOR : ALIAS FOR N7[60];
   TK24_PUMP : ALIAS FOR N7[80];
   TK25_COLOR : ALIAS FOR N7[61];
   TK25_PUMP : ALIAS FOR N7[81];
   TK26_COLOR : ALIAS FOR N7[62];
   TK26_PUMP : ALIAS FOR N7[82];
   tmrSetWaterOil : TIMER := (PRE := 1000);
   Toss_Bit : BOOL := 1;
   tpCreateTicket : BOOL;
   tpCreateTicketRecvd : DINT;
   tpLocation : DINT := 1;
   tpNewGrossWt : BOOL;
   tpNewGrossWtRecvd : DINT;
   tpNewGrossWtSent : BOOL;
   tpNewTareWt : BOOL;
   tpNewTareWtRecvd : DINT;
   tpNewTareWtSent : BOOL;
   tpShowGrossPB : BOOL;
   tpShowTarePB : BOOL;
   tpVarsTrtsComplete : BOOL;
   Treat_Produced : DINT; {produced}
   Treater_Remote_In : DINT;
   Treater_Remote_Out : DINT := 2; {produced}
   TRT_ARRAY : STRING[50] := ([1] := '99999 - Water', [2] := '28022 - Albaugh NWGG .25', [3] := '28031 - Evergol Energy', [4] := '28060 - Macho 600ST', [5] := '28050 - Vibrance Extreme Bulk', [6] := '28122 - Cruiser Maxx High Residue .33', [7] := '28080 - TBZ', [8] := '29140 - Wuxal Terios', [9] := '12000 - Blue Dye', [10] := '99998 - Oil', [11] := '28100 - Apron', [12] := '28085 - Stamina Treat');
   TRT_CNT : DINT;
   TRT_CNT_ONS : DINT;
   Trt_CntStore : DINT := 2;
   TRT_PumpRATE : DINT[50] := ([1] := 80, [2] := 43, [3] := 35, [4] := 30, [5] := 29, [6] := 30, [7] := 30, [8] := 40, [10] := 22);
   TRT_PumpTotOz : DINT[50];
   TRT_TICKETtable : STRING[100] := ([0] := 'Empty', [1] := 'Empty', [2] := 'Empty', [3] := 'Empty', [4] := 'Empty', [5] := 'Empty', [6] := 'Empty', [7] := 'Empty', [8] := '28100 - Apron', [9] := '28085 - Stamina Treat', [10] := '28122 - Cruiser Maxx High Residue .33', [11] := '28050 - Vibrance Extreme Bulk');
   TRT_TickettableItemNo : DINT[50];
   TRT_TICKETtableRate : DINT[100];
   TRT_TICKETtableTotalOz : DINT[100];
   TrtTrimTemp : STRING := '28022 ';
   Truck_Scales : udt_Truck_Scale[2] := ([0].Rate_Stable := 1, [0].Rate_Tol := 1.0, [1].Rate_Tol := 1.0, [1].Faulted := 1, [1].Int_Rate := -15872);
   VAR_CNT : DINT;
   VAR_CNT_ONS : DINT := 1;
   Var_CntStore : DINT := 1;
   var_control : CONTROL;
   var_control1 : CONTROL;
   VAR_TICKETtable : STRING[20] := ([0] := 'Empty', [1] := 'Empty', [2] := 'Empty', [3] := 'Empty', [4] := 'Empty', [5] := 'Empty', [6] := 'Empty', [7] := 'Empty', [8] := 'Empty', [9] := 'Empty', [10] := 'Empty', [11] := 'Empty', [12] := 'Empty', [13] := 'Empty', [14] := 'Empty', [15] := 'Empty', [16] := 'Empty', [17] := 'Empty', [18] := 'Empty', [19] := 'Empty');
   VAR_TickettableItemNo : DINT[50];
   VAR_TICKETtableRate : DINT[100];
   VAR_TICKETtableWt : DINT[100];
   Varieties : Variety[1000] := ([0].Name := 'ALUM', [0].Class := 'Certified', [1].Name := 'ALUM', [1].Class := 'Common', [2].Name := 'ALUM', [2].Class := 'Foundation', [3].Name := 'ALUM', [3].Class := 'Registered', [4].Name := 'AP 700', [4].Class := 'Certified', [5].Name := 'AP 700', [5].Class := 'Common', [6].Name := 'AP 700', [6].Class := 'Foundation', [7].Name := 'AP 700', [7].Class := 'Registered', [8].Name := 'Aragorn', [8].Class := 'Certified', [9].Name := 'Aragorn', [9].Class := 'Common', [10].Name := 'Aragorn', [10].Class := 'Foundation', [11].Name := 'Aragorn', [11].Class := 'Registered', [12].Name := 'Aragorn-Spokane Seed', [12].Class := 'Certified', [13].Name := 'Aragorn-Spokane Seed', [13].Class := 'Common', [14].Name := 'Aragorn-Spokane Seed', [14].Class := 'Foundation', [15].Name := 'Aragorn-Spokane Seed', [15].Class := 'Registered', [16].Name := 'Aragorn-Spokane Seed-Day', [16].Class := 'Certified', [17].Name := 'Aragorn-Spokane Seed-Day', [17].Class := 'Common', [18].Name := 'Aragorn-Spokane Seed-Day', [18].Class := 'Foundation', [19].Name := 'Aragorn-Spokane Seed-Day', [19].Class := 'Registered', [20].Name := 'Ariel', [20].Class := 'Certified', [21].Name := 'Ariel', [21].Class := 'Common', [22].Name := 'Ariel', [22].Class := 'Foundation', [23].Name := 'Ariel', [23].Class := 'Registered', [24].Name := 'ArtDeco', [24].Class := 'Certified', [25].Name := 'ArtDeco', [25].Class := 'Common', [26].Name := 'ArtDeco', [26].Class := 'Foundation', [27].Name := 'ArtDeco', [27].Class := 'Registered', [28].Name := 'Azimut', [28].Class := 'Certified', [29].Name := 'Azimut', [29].Class := 'Common',
        [30].Name := 'Azimut', [30].Class := 'Foundation', [31].Name := 'Azimut', [31].Class := 'Registered', [32].Name := 'Babe ', [32].Class := 'Certified', [33].Name := 'Babe ', [33].Class := 'Common', [34].Name := 'Babe ', [34].Class := 'Foundation', [35].Name := 'Babe ', [35].Class := 'Registered', [36].Name := 'Banner-Anderson', [36].Class := 'Certified', [37].Name := 'Banner-Anderson', [37].Class := 'Common', [38].Name := 'Banner-Anderson', [38].Class := 'Foundation', [39].Name := 'Banner-Anderson', [39].Class := 'Registered', [40].Name := 'Banner-Anderson-Day', [40].Class := 'Certified', [41].Name := 'Banner-Anderson-Day', [41].Class := 'Common', [42].Name := 'Banner-Anderson-Day', [42].Class := 'Foundation', [43].Name := 'Banner-Anderson-Day', [43].Class := 'Registered', [44].Name := 'Banner-Columbia Grain', [44].Class := 'Certified', [45].Name := 'Banner-Columbia Grain', [45].Class := 'Common', [46].Name := 'Banner-Columbia Grain', [46].Class := 'Foundation', [47].Name := 'Banner-Columbia Grain', [47].Class := 'Registered', [48].Name := 'Banner-Columbian Grian-Day', [48].Class := 'Certified', [49].Name := 'Banner-Columbian Grian-Day', [49].Class := 'Common', [50].Name := 'Banner-Columbian Grian-Day', [50].Class := 'Foundation', [51].Name := 'Banner-Columbian Grian-Day', [51].Class := 'Registered', [52].Name := 'Banner-PNWFC', [52].Class := 'Certified', [53].Name := 'Banner-PNWFC', [53].Class := 'Common', [54].Name := 'Banner-PNWFC', [54].Class := 'Foundation', [55].Name := 'Banner-PNWFC', [55].Class := 'Registered', [56].Name := 'Biancor', [56].Class := 'Certified', [57].Name := 'Biancor', [57].Class := 'Common', [58].Name := 'Biancor', [58].Class := 'Foundation', [59].Name := 'Biancor', [59].Class := 'Registered',
        [60].Name := 'Billy Beans PNWFC', [60].Class := 'Certified', [61].Name := 'Billy Beans PNWFC', [61].Class := 'Common', [62].Name := 'Billy Beans PNWFC', [62].Class := 'Foundation', [63].Name := 'Billy Beans PNWFC', [63].Class := 'Registered', [64].Name := 'Bobtail', [64].Class := 'Certified', [65].Name := 'Bobtail', [65].Class := 'Common', [66].Name := 'Bobtail', [66].Class := 'Foundation', [67].Name := 'Bobtail', [67].Class := 'Registered', [68].Name := 'Brawl', [68].Class := 'Certified', [69].Name := 'Brawl', [69].Class := 'Common', [70].Name := 'Brawl', [70].Class := 'Foundation', [71].Name := 'Brawl', [71].Class := 'Registered', [72].Name := 'Brundage', [72].Class := 'Certified', [73].Name := 'Brundage', [73].Class := 'Common', [74].Name := 'Brundage', [74].Class := 'Foundation', [75].Name := 'Brundage', [75].Class := 'Registered', [76].Name := 'Buck Pronto', [76].Class := 'Certified', [77].Name := 'Buck Pronto', [77].Class := 'Common', [78].Name := 'Buck Pronto', [78].Class := 'Foundation', [79].Name := 'Buck Pronto', [79].Class := 'Registered', [80].Name := 'Cara Club', [80].Class := 'Certified', [81].Name := 'Cara Club', [81].Class := 'Common', [82].Name := 'Cara Club', [82].Class := 'Foundation', [83].Name := 'Cara Club', [83].Class := 'Registered', [84].Name := 'Chet', [84].Class := 'Certified', [85].Name := 'Chet', [85].Class := 'Common', [86].Name := 'Chet', [86].Class := 'Foundation', [87].Name := 'Chet', [87].Class := 'Registered', [88].Name := 'Clearstone', [88].Class := 'Certified', [89].Name := 'Clearstone', [89].Class := 'Common',
        [90].Name := 'Clearstone', [90].Class := 'Foundation', [91].Name := 'Clearstone', [91].Class := 'Registered', [92].Name := 'Coda Club', [92].Class := 'Certified', [93].Name := 'Coda Club', [93].Class := 'Common', [94].Name := 'Coda Club', [94].Class := 'Foundation', [95].Name := 'Coda Club', [95].Class := 'Registered', [96].Name := 'Colonia', [96].Class := 'Certified', [97].Name := 'Colonia', [97].Class := 'Common', [98].Name := 'Colonia', [98].Class := 'Foundation', [99].Name := 'Colonia', [99].Class := 'Registered', [100].Name := 'Columbian', [100].Class := 'Certified', [101].Name := 'Columbian', [101].Class := 'Common', [102].Name := 'Columbian', [102].Class := 'Foundation', [103].Name := 'Columbian', [103].Class := 'Registered', [104].Name := 'Columbian Spokane Seed', [104].Class := 'Certified', [105].Name := 'Columbian Spokane Seed', [105].Class := 'Common', [106].Name := 'Columbian Spokane Seed', [106].Class := 'Foundation', [107].Name := 'Columbian Spokane Seed', [107].Class := 'Registered', [108].Name := 'Columbian Spokane Seed-Day', [108].Class := 'Certified', [109].Name := 'Columbian Spokane Seed-Day', [109].Class := 'Common', [110].Name := 'Columbian Spokane Seed-Day', [110].Class := 'Foundation', [111].Name := 'Columbian Spokane Seed-Day', [111].Class := 'Registered', [112].Name := 'Diva Spring', [112].Class := 'Certified', [113].Name := 'Diva Spring', [113].Class := 'Common', [114].Name := 'Diva Spring', [114].Class := 'Foundation', [115].Name := 'Diva Spring', [115].Class := 'Registered', [116].Name := 'Drive (7105)', [116].Class := 'Certified', [117].Name := 'Drive (7105)', [117].Class := 'Common', [118].Name := 'Drive (7105)', [118].Class := 'Foundation', [119].Name := 'Drive (7105)', [119].Class := 'Registered',
        [120].Name := 'Expresso', [120].Class := 'Certified', [121].Name := 'Expresso', [121].Class := 'Common', [122].Name := 'Expresso', [122].Class := 'Foundation', [123].Name := 'Expresso', [123].Class := 'Registered', [124].Name := 'Frontier', [124].Class := 'Certified', [125].Name := 'Frontier', [125].Class := 'Common', [126].Name := 'Frontier', [126].Class := 'Foundation', [127].Name := 'Frontier', [127].Class := 'Registered', [128].Name := 'Genie', [128].Class := 'Certified', [129].Name := 'Genie', [129].Class := 'Common', [130].Name := 'Genie', [130].Class := 'Foundation', [131].Name := 'Genie', [131].Class := 'Registered', [132].Name := 'Ginny-Spokane Seed', [132].Class := 'Certified', [133].Name := 'Ginny-Spokane Seed', [133].Class := 'Common', [134].Name := 'Ginny-Spokane Seed', [134].Class := 'Foundation', [135].Name := 'Ginny-Spokane Seed', [135].Class := 'Registered', [136].Name := 'Glee ', [136].Class := 'Certified', [137].Name := 'Glee ', [137].Class := 'Common', [138].Name := 'Glee ', [138].Class := 'Foundation', [139].Name := 'Glee ', [139].Class := 'Registered', [140].Name := 'Hard White Wheat', [140].Class := 'Certified', [141].Name := 'Hard White Wheat', [141].Class := 'Common', [142].Name := 'Hard White Wheat', [142].Class := 'Foundation', [143].Name := 'Hard White Wheat', [143].Class := 'Registered', [144].Name := 'Haybet', [144].Class := 'Certified', [145].Name := 'Haybet', [145].Class := 'Common', [146].Name := 'Haybet', [146].Class := 'Foundation', [147].Name := 'Haybet', [147].Class := 'Registered', [148].Name := 'Huffman', [148].Class := 'Certified', [149].Name := 'Huffman', [149].Class := 'Common',
        [150].Name := 'Huffman', [150].Class := 'Foundation', [151].Name := 'Huffman', [151].Class := 'Registered', [152].Name := 'Iron', [152].Class := 'Certified', [153].Name := 'Iron', [153].Class := 'Common', [154].Name := 'Iron', [154].Class := 'Foundation', [155].Name := 'Iron', [155].Class := 'Registered', [156].Name := 'Jasper', [156].Class := 'Certified', [157].Name := 'Jasper', [157].Class := 'Common', [158].Name := 'Jasper', [158].Class := 'Foundation', [159].Name := 'Jasper', [159].Class := 'Registered', [160].Name := 'JD Club Spring', [160].Class := 'Certified', [161].Name := 'JD Club Spring', [161].Class := 'Common', [162].Name := 'JD Club Spring', [162].Class := 'Foundation', [163].Name := 'JD Club Spring', [163].Class := 'Registered', [164].Name := 'Jefferson', [164].Class := 'Certified', [165].Name := 'Jefferson', [165].Class := 'Common', [166].Name := 'Jefferson', [166].Class := 'Foundation', [167].Name := 'Jefferson', [167].Class := 'Registered', [168].Name := 'Jet', [168].Class := 'Certified', [169].Name := 'Jet', [169].Class := 'Common', [170].Name := 'Jet', [170].Class := 'Foundation', [171].Name := 'Jet', [171].Class := 'Registered', [172].Name := 'Kaseberg', [172].Class := 'Certified', [173].Name := 'Kaseberg', [173].Class := 'Common', [174].Name := 'Kaseberg', [174].Class := 'Foundation', [175].Name := 'Kaseberg', [175].Class := 'Registered', [176].Name := 'Keldin ', [176].Class := 'Certified', [177].Name := 'Keldin ', [177].Class := 'Common', [178].Name := 'Keldin ', [178].Class := 'Foundation', [179].Name := 'Keldin ', [179].Class := 'Registered',
        [180].Name := 'Kelse', [180].Class := 'Certified', [181].Name := 'Kelse', [181].Class := 'Common', [182].Name := 'Kelse', [182].Class := 'Foundation', [183].Name := 'Kelse', [183].Class := 'Registered', [184].Name := 'Latah', [184].Class := 'Certified', [185].Name := 'Latah', [185].Class := 'Common', [186].Name := 'Latah', [186].Class := 'Foundation', [187].Name := 'Latah', [187].Class := 'Registered', [188].Name := 'Lenetah', [188].Class := 'Certified', [189].Name := 'Lenetah', [189].Class := 'Common', [190].Name := 'Lenetah', [190].Class := 'Foundation', [191].Name := 'Lenetah', [191].Class := 'Registered', [192].Name := 'Levina', [192].Class := 'Certified', [193].Name := 'Levina', [193].Class := 'Common', [194].Name := 'Levina', [194].Class := 'Foundation', [195].Name := 'Levina', [195].Class := 'Registered', [196].Name := 'Louise Spring', [196].Class := 'Certified', [197].Name := 'Louise Spring', [197].Class := 'Common', [198].Name := 'Louise Spring', [198].Class := 'Foundation', [199].Name := 'Louise Spring', [199].Class := 'Registered', [200].Name := 'Madsen', [200].Class := 'Certified', [201].Name := 'Madsen', [201].Class := 'Common', [202].Name := 'Madsen', [202].Class := 'Foundation', [203].Name := 'Madsen', [203].Class := 'Registered', [204].Name := 'Majic', [204].Class := 'Certified', [205].Name := 'Majic', [205].Class := 'Common', [206].Name := 'Majic', [206].Class := 'Foundation', [207].Name := 'Majic', [207].Class := 'Registered', [208].Name := 'Mary', [208].Class := 'Certified', [209].Name := 'Mary', [209].Class := 'Common',
        [210].Name := 'Mary', [210].Class := 'Foundation', [211].Name := 'Mary', [211].Class := 'Registered', [212].Name := 'Northwest Tandem', [212].Class := 'Certified', [213].Name := 'Northwest Tandem', [213].Class := 'Common', [214].Name := 'Northwest Tandem', [214].Class := 'Foundation', [215].Name := 'Northwest Tandem', [215].Class := 'Registered', [216].Name := 'NW Duet', [216].Class := 'Certified', [217].Name := 'NW Duet', [217].Class := 'Common', [218].Name := 'NW Duet', [218].Class := 'Foundation', [219].Name := 'NW Duet', [219].Class := 'Registered', [220].Name := 'ORCF 101', [220].Class := 'Certified', [221].Name := 'ORCF 101', [221].Class := 'Common', [222].Name := 'ORCF 101', [222].Class := 'Foundation', [223].Name := 'ORCF 101', [223].Class := 'Registered', [224].Name := 'ORCF 102', [224].Class := 'Certified', [225].Name := 'ORCF 102', [225].Class := 'Common', [226].Name := 'ORCF 102', [226].Class := 'Foundation', [227].Name := 'ORCF 102', [227].Class := 'Registered', [228].Name := 'Ovation', [228].Class := 'Certified', [229].Name := 'Ovation', [229].Class := 'Common', [230].Name := 'Ovation', [230].Class := 'Foundation', [231].Name := 'Ovation', [231].Class := 'Registered', [232].Name := 'Palouse', [232].Class := 'Certified', [233].Name := 'Palouse', [233].Class := 'Common', [234].Name := 'Palouse', [234].Class := 'Foundation', [235].Name := 'Palouse', [235].Class := 'Registered', [236].Name := 'Puma', [236].Class := 'Certified', [237].Name := 'Puma', [237].Class := 'Common', [238].Name := 'Puma', [238].Class := 'Foundation', [239].Name := 'Puma', [239].Class := 'Registered',
        [240].Name := 'Rod', [240].Class := 'Certified', [241].Name := 'Rod', [241].Class := 'Common', [242].Name := 'Rod', [242].Class := 'Foundation', [243].Name := 'Rod', [243].Class := 'Registered', [244].Name := 'Scotch-Spokane Seed', [244].Class := 'Certified', [245].Name := 'Scotch-Spokane Seed', [245].Class := 'Common', [246].Name := 'Scotch-Spokane Seed', [246].Class := 'Foundation', [247].Name := 'Scotch-Spokane Seed', [247].Class := 'Registered', [248].Name := 'Scotch-Spokane Seed-Day', [248].Class := 'Certified', [249].Name := 'Scotch-Spokane Seed-Day', [249].Class := 'Common', [250].Name := 'Scotch-Spokane Seed-Day', [250].Class := 'Foundation', [251].Name := 'Scotch-Spokane Seed-Day', [251].Class := 'Registered', [252].Name := 'Seahawk', [252].Class := 'Certified', [253].Name := 'Seahawk', [253].Class := 'Common', [254].Name := 'Seahawk', [254].Class := 'Foundation', [255].Name := 'Seahawk', [255].Class := 'Registered', [256].Name := 'Sierra', [256].Class := 'Certified', [257].Name := 'Sierra', [257].Class := 'Common', [258].Name := 'Sierra', [258].Class := 'Foundation', [259].Name := 'Sierra', [259].Class := 'Registered', [260].Name := 'Sierra PNWFC', [260].Class := 'Certified', [261].Name := 'Sierra PNWFC', [261].Class := 'Common', [262].Name := 'Sierra PNWFC', [262].Class := 'Foundation', [263].Name := 'Sierra PNWFC', [263].Class := 'Registered', [264].Name := 'Sierra Spokane Seed', [264].Class := 'Certified', [265].Name := 'Sierra Spokane Seed', [265].Class := 'Common', [266].Name := 'Sierra Spokane Seed', [266].Class := 'Foundation', [267].Name := 'Sierra Spokane Seed', [267].Class := 'Registered', [268].Name := 'Skiles', [268].Class := 'Certified', [269].Name := 'Skiles', [269].Class := 'Common',
        [270].Name := 'Skiles', [270].Class := 'Foundation', [271].Name := 'Skiles', [271].Class := 'Registered', [272].Name := 'Solano', [272].Class := 'Certified', [273].Name := 'Solano', [273].Class := 'Common', [274].Name := 'Solano', [274].Class := 'Foundation', [275].Name := 'Solano', [275].Class := 'Registered', [276].Name := 'Stephens', [276].Class := 'Certified', [277].Name := 'Stephens', [277].Class := 'Common', [278].Name := 'Stephens', [278].Class := 'Foundation', [279].Name := 'Stephens', [279].Class := 'Registered', [280].Name := 'Sy 107', [280].Class := 'Certified', [281].Name := 'Sy 107', [281].Class := 'Common', [282].Name := 'Sy 107', [282].Class := 'Foundation', [283].Name := 'Sy 107', [283].Class := 'Registered', [284].Name := 'SY 605', [284].Class := 'Certified', [285].Name := 'SY 605', [285].Class := 'Common', [286].Name := 'SY 605', [286].Class := 'Foundation', [287].Name := 'SY 605', [287].Class := 'Registered', [288].Name := 'SY Assure', [288].Class := 'Certified', [289].Name := 'SY Assure', [289].Class := 'Common', [290].Name := 'SY Assure', [290].Class := 'Foundation', [291].Name := 'SY Assure', [291].Class := 'Registered', [292].Name := 'Test', [292].Class := 'Certified', [293].Name := 'Test', [293].Class := 'Common', [294].Name := 'Test', [294].Class := 'Foundation', [295].Name := 'Test', [295].Class := 'Registered', [296].Name := 'Tubbs', [296].Class := 'Certified', [297].Name := 'Tubbs', [297].Class := 'Common', [298].Name := 'Tubbs', [298].Class := 'Foundation', [299].Name := 'Tubbs', [299].Class := 'Registered',
        [300].Name := 'Universal-Spokane Seed', [300].Class := 'Certified', [301].Name := 'Universal-Spokane Seed', [301].Class := 'Common', [302].Name := 'Universal-Spokane Seed', [302].Class := 'Foundation', [303].Name := 'Universal-Spokane Seed', [303].Class := 'Registered', [304].Name := 'Vespa', [304].Class := 'Certified', [305].Name := 'Vespa', [305].Class := 'Common', [306].Name := 'Vespa', [306].Class := 'Foundation', [307].Name := 'Vespa', [307].Class := 'Registered', [308].Name := 'WB 1035 CL spring', [308].Class := 'Certified', [309].Name := 'WB 1035 CL spring', [309].Class := 'Common', [310].Name := 'WB 1035 CL spring', [310].Class := 'Foundation', [311].Name := 'WB 1035 CL spring', [311].Class := 'Registered', [312].Name := 'WB 1070', [312].Class := 'Certified', [313].Name := 'WB 1070', [313].Class := 'Common', [314].Name := 'WB 1070', [314].Class := 'Foundation', [315].Name := 'WB 1070', [315].Class := 'Registered', [316].Name := 'WB 1376', [316].Class := 'Certified', [317].Name := 'WB 1376', [317].Class := 'Common', [318].Name := 'WB 1376', [318].Class := 'Foundation', [319].Name := 'WB 1376', [319].Class := 'Registered', [320].Name := 'WB 1529', [320].Class := 'Certified', [321].Name := 'WB 1529', [321].Class := 'Common', [322].Name := 'WB 1529', [322].Class := 'Foundation', [323].Name := 'WB 1529', [323].Class := 'Registered', [324].Name := 'WB 1604', [324].Class := 'Certified', [325].Name := 'WB 1604', [325].Class := 'Common', [326].Name := 'WB 1604', [326].Class := 'Foundation', [327].Name := 'WB 1604', [327].Class := 'Registered', [328].Name := 'WB 528', [328].Class := 'Certified', [329].Name := 'WB 528', [329].Class := 'Common',
        [330].Name := 'WB 528', [330].Class := 'Foundation', [331].Name := 'WB 528', [331].Class := 'Registered', [332].Name := 'WB 6121 spring', [332].Class := 'Certified', [333].Name := 'WB 6121 spring', [333].Class := 'Common', [334].Name := 'WB 6121 spring', [334].Class := 'Foundation', [335].Name := 'WB 6121 spring', [335].Class := 'Registered', [336].Name := 'WB 6341 Spring', [336].Class := 'Certified', [337].Name := 'WB 6341 Spring', [337].Class := 'Common', [338].Name := 'WB 6341 Spring', [338].Class := 'Foundation', [339].Name := 'WB 6341 Spring', [339].Class := 'Registered', [340].Name := 'WB 9411', [340].Class := 'Certified', [341].Name := 'WB 9411', [341].Class := 'Common', [342].Name := 'WB 9411', [342].Class := 'Foundation', [343].Name := 'WB 9411', [343].Class := 'Registered', [344].Name := 'WB 9518', [344].Class := 'Certified', [345].Name := 'WB 9518', [345].Class := 'Common', [346].Name := 'WB 9518', [346].Class := 'Foundation', [347].Name := 'WB 9518', [347].Class := 'Registered', [348].Name := 'WB523', [348].Class := 'Certified', [349].Name := 'WB523', [349].Class := 'Common', [350].Name := 'WB523', [350].Class := 'Foundation', [351].Name := 'WB523', [351].Class := 'Registered', [352].Name := 'Xerpha', [352].Class := 'Certified', [353].Name := 'Xerpha', [353].Class := 'Common', [354].Name := 'Xerpha', [354].Class := 'Foundation', [355].Name := 'Xerpha', [355].Class := 'Registered');
   varIndx : DINT;
   vartableONS : DINT := 3;
   VarTrimTemp : STRING := '843001';
   VIRTUAL_BT : ALIAS FOR N20[5].13;
   VIRTUAL_BT1 : ALIAS FOR N23[0].12;
   VIRTUAL_BT2 : ALIAS FOR N23[0].13;
   zzzRealtmp : REAL := 30.73328;
   zzzsqlVaritiesRevd : BOOL;
   zzztmpSqlDataArryDINT : DINT[10];
   zzztmpSqlDataArryFLT : REAL[10];
   zzztmpSqlDataDINT : DINT := 1000;
   zzztmpSqlDataFLT : REAL;
   zzztmpSqlDataSTR : STRING;
   zzztmpTANKtest : DINT[10];
   zzzz_22_GATE_PO_STOR : DINT;
   zzzzProcessAll : DINT;
   zzzzSTRING : STRING := '821001 ArtDeco SWW';
   zzzzTestGrossWt : BOOL;
   zzzzTestTareWt : BOOL;
   zzzztmpDINT : DINT[10];
   zzzzVAR_CNT_ONS : BOOL;
   zzzzzTestBit : BOOL;
END_VAR

PROGRAM _2_MAIN   (* main routine _02_MAIN *)
VAR
   Flow_Gal2Oz : FBD_MATH := (SourceB := 0.015);
   GRT_01 : FBD_COMPARE := (SourceB := 75.0);
   HOUR_METERS : DINT;
   LES_01 : FBD_COMPARE;
   LES_02 : FBD_COMPARE;
   SCL_01 : SCALE := (InRawMax := 100.0, InEUMax := 4000.0);
   SCL_02 : SCALE := (In := 28776.0, InRawMin := 31000.0, InEUMax := 3200.0, Status := 16#0000_0003, InstructFault := 1, InRawRangeInv := 1);
   SCL_03 : SCALE := (In := 6569.0, InRawMax := 13975.0, InRawMin := 578.0, InEUMax := 3000.0, Out := 1341.569);
   SCL_04 : SCALE;
   SCL_05 : SCALE;
   SCL_06 : SCALE := (InRawMax := 60.0, InEUMax := 32767.0);
   SCL_07 : SCALE := (In := 46.0, InRawMax := 60.0, InEUMax := 31000.0, Out := 23766.668);
   SCL_08 : SCALE := (In := 48.0, InRawMax := 60.0, InEUMax := 31000.0, Out := 24800.0);
   SCL_09 : SCALE := (In := 53.0, InRawMax := 60.0, InEUMax := 31000.0, Out := 27383.334);
   SEL_01 : SELECT;
   SUB_01 : FBD_MATH;
   Test_Bit : BOOL;
   TOT_01 : TOTALIZER := (Gain := 1.0, ProgProgReq := 1, ProgStartReq := 1, RTSTime := 1, Total := 3307.86, OldTotal := 877.80005, ProgOper := 1, RunStop := 1, TargetFlag := 1, TargetDev1Flag := 1, TargetDev2Flag := 1, LowInCutoffFlag := 1, DeltaT := 0.004);
END_VAR

ROUTINE _02_MAIN   (* ladder *)
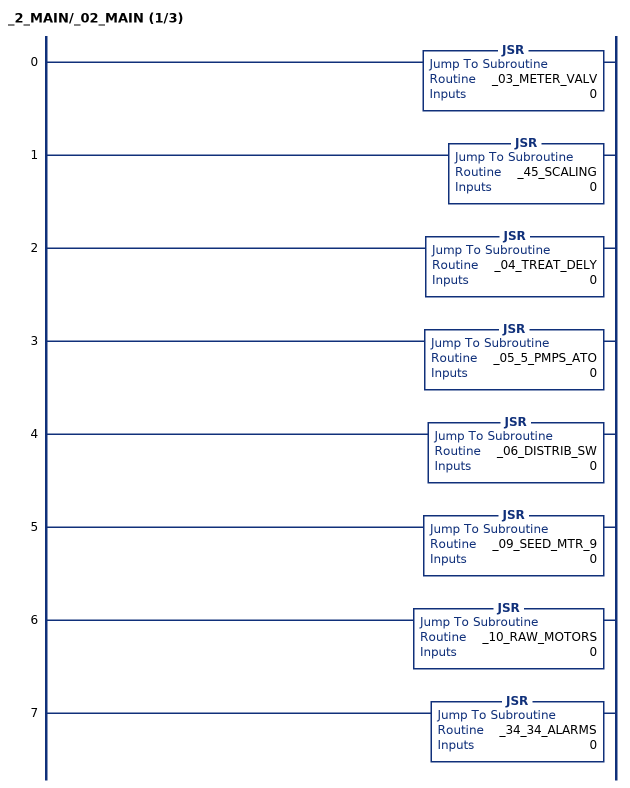
   0: JSR(_03_METER_VALV,0);
   1: JSR(_45_SCALING,0);
   2: JSR(_04_TREAT_DELY,0);
   3: JSR(_05_5_PMPS_ATO,0);
   4: JSR(_06_DISTRIB_SW,0);
   5: JSR(_09_SEED_MTR_9,0);
   6: JSR(_10_RAW_MOTORS,0);
   7: JSR(_34_34_ALARMS,0);
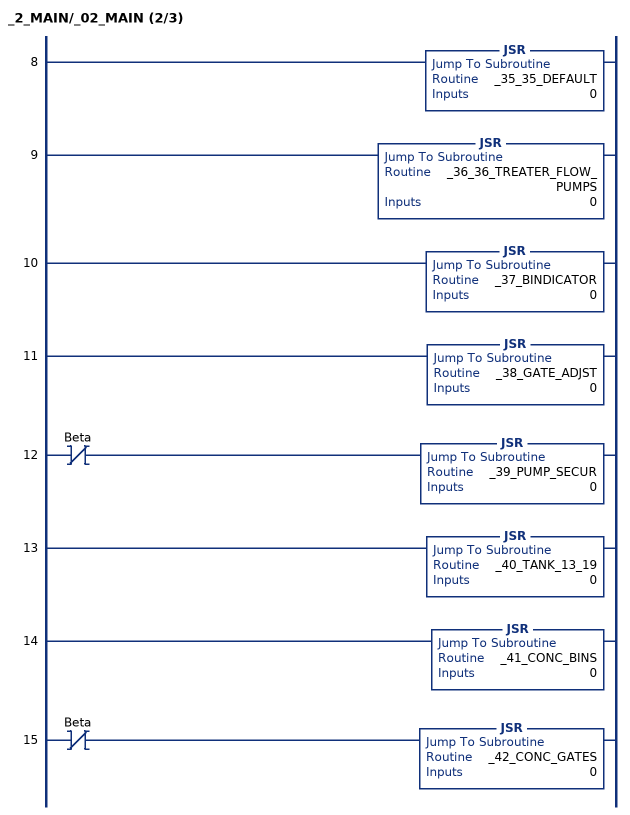
   8: JSR(_35_35_DEFAULT,0);
   9: JSR(_36_36_TREATER_FLOW_PUMPS,0);
   10: JSR(_37_BINDICATOR,0);
   11: JSR(_38_GATE_ADJST,0);
   12: XIO(Beta)JSR(_39_PUMP_SECUR,0);
   13: JSR(_40_TANK_13_19,0);
   14: JSR(_41_CONC_BINS,0);
   15: XIO(Beta)JSR(_42_CONC_GATES,0);
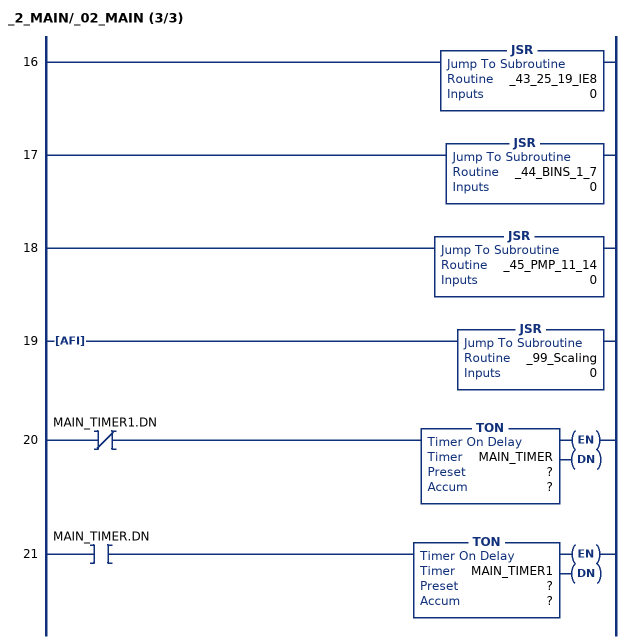
   16: JSR(_43_25_19_IE8,0);
   17: JSR(_44_BINS_1_7,0);
   18: JSR(_45_PMP_11_14,0);
   19: AFI()JSR(_99_Scaling,0);
   20: XIO(MAIN_TIMER1.DN)TON(MAIN_TIMER,?,?);
   21: XIC(MAIN_TIMER.DN)TON(MAIN_TIMER1,?,?);
END_ROUTINE

ROUTINE _03_METER_VALV   (* ladder *)
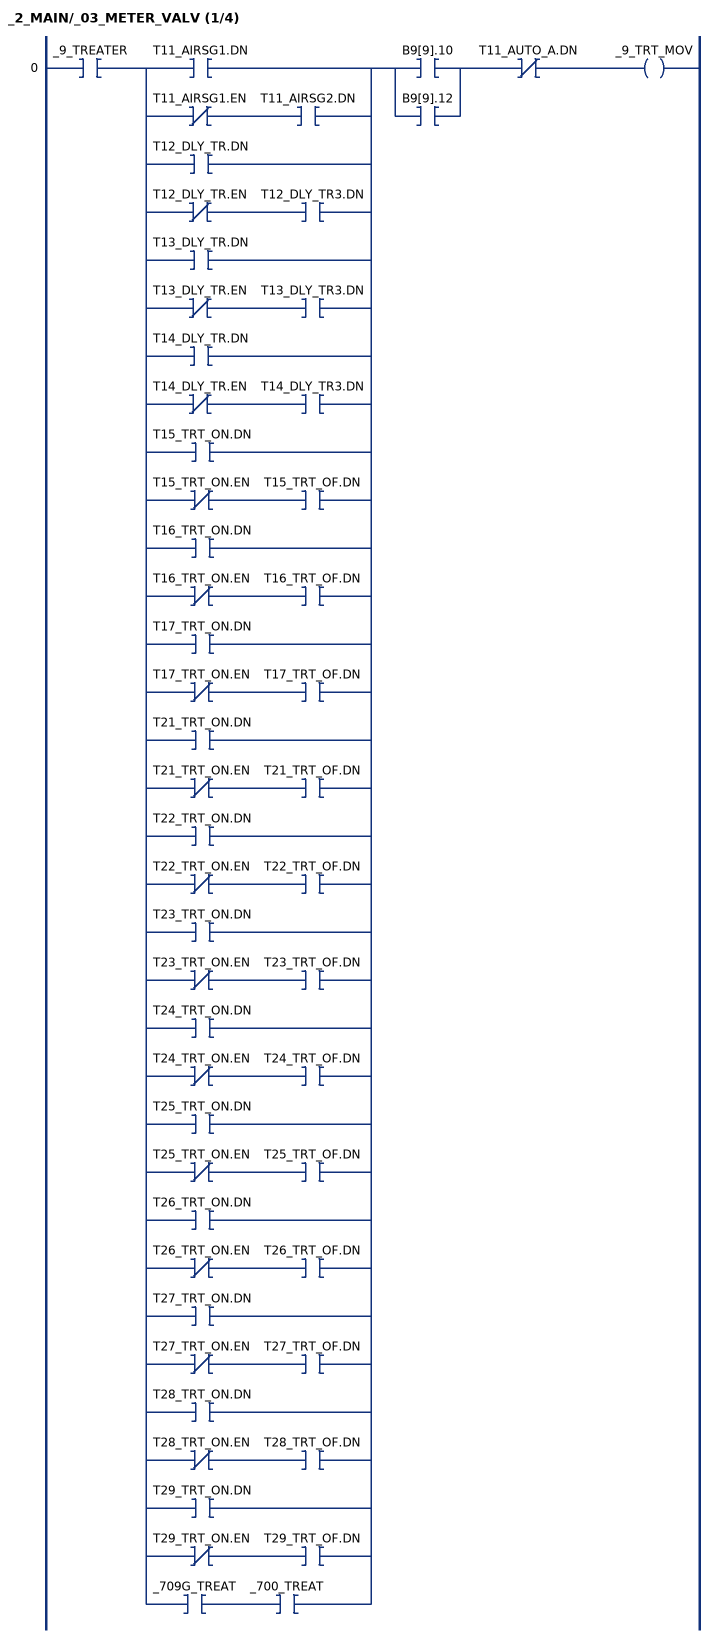
   0: XIC(_9_TREATER)[XIC(T11_AIRSG1.DN) ,XIO(T11_AIRSG1.EN) XIC(T11_AIRSG2.DN) ,XIC(T12_DLY_TR.DN) ,XIO(T12_DLY_TR.EN) XIC(T12_DLY_TR3.DN) ,XIC(T13_DLY_TR.DN) ,XIO(T13_DLY_TR.EN) XIC(T13_DLY_TR3.DN) ,XIC(T14_DLY_TR.DN) ,XIO(T14_DLY_TR.EN) XIC(T14_DLY_TR3.DN) ,XIC(T15_TRT_ON.DN) ,XIO(T15_TRT_ON.EN) XIC(T15_TRT_OF.DN) ,XIC(T16_TRT_ON.DN) ,XIO(T16_TRT_ON.EN) XIC(T16_TRT_OF.DN) ,XIC(T17_TRT_ON.DN) ,XIO(T17_TRT_ON.EN) XIC(T17_TRT_OF.DN) ,XIC(T21_TRT_ON.DN) ,XIO(T21_TRT_ON.EN) XIC(T21_TRT_OF.DN) ,XIC(T22_TRT_ON.DN) ,XIO(T22_TRT_ON.EN) XIC(T22_TRT_OF.DN) ,XIC(T23_TRT_ON.DN) ,XIO(T23_TRT_ON.EN) XIC(T23_TRT_OF.DN) ,XIC(T24_TRT_ON.DN) ,XIO(T24_TRT_ON.EN) XIC(T24_TRT_OF.DN) ,XIC(T25_TRT_ON.DN) ,XIO(T25_TRT_ON.EN) XIC(T25_TRT_OF.DN) ,XIC(T26_TRT_ON.DN) ,XIO(T26_TRT_ON.EN) XIC(T26_TRT_OF.DN) ,XIC(T27_TRT_ON.DN) ,XIO(T27_TRT_ON.EN) XIC(T27_TRT_OF.DN) ,XIC(T28_TRT_ON.DN) ,XIO(T28_TRT_ON.EN) XIC(T28_TRT_OF.DN) ,XIC(T29_TRT_ON.DN) ,XIO(T29_TRT_ON.EN) XIC(T29_TRT_OF.DN) ,XIC(_709G_TREAT) XIC(_700_TREAT) ][XIC(B9[9].10) ,XIC(B9[9].12) ]XIO(T11_AUTO_A.DN)OTE(_9_TRT_MOV);
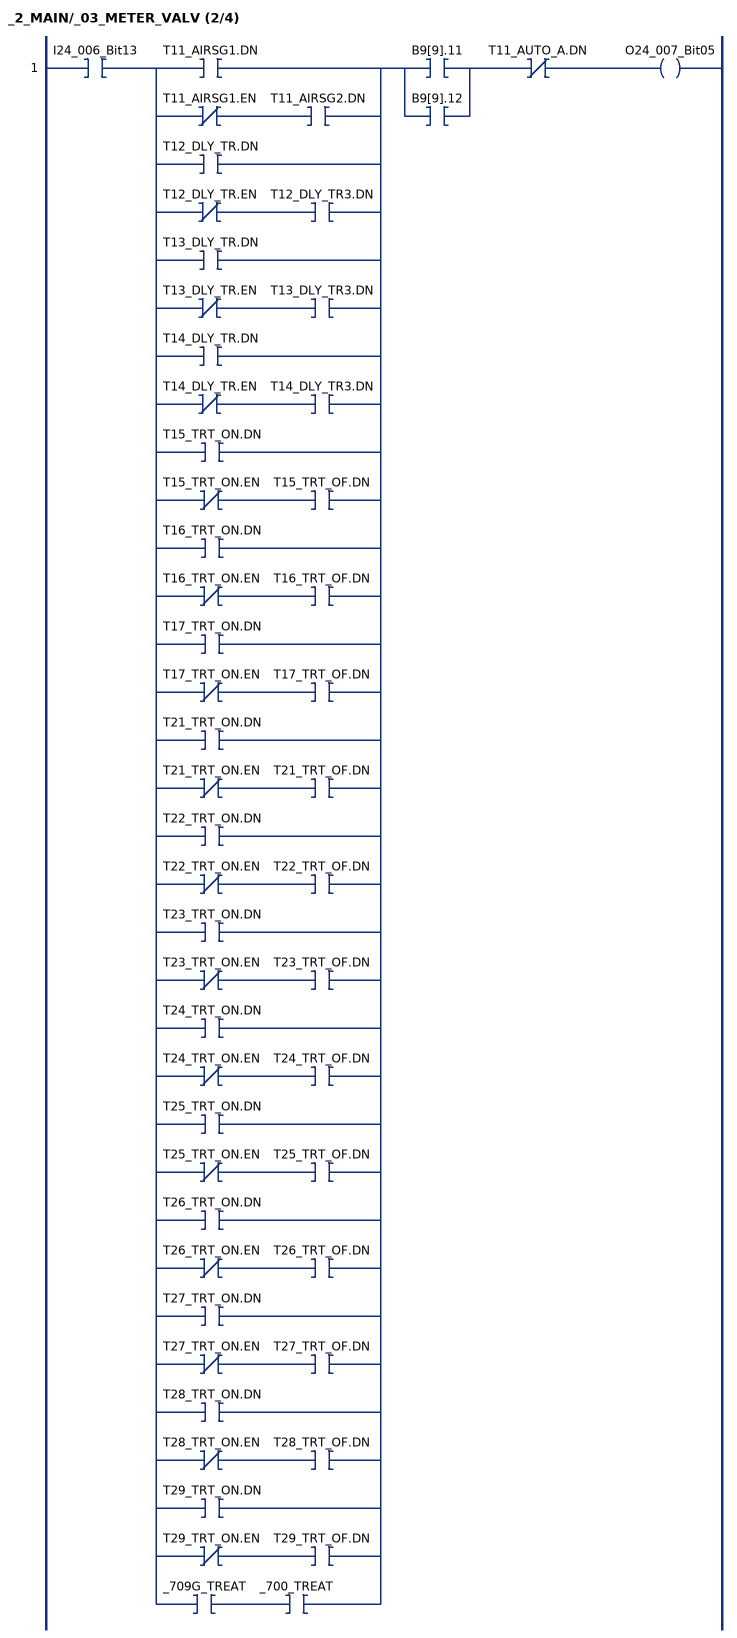
   1: XIC(I24_006_Bit13)[XIC(T11_AIRSG1.DN) ,XIO(T11_AIRSG1.EN) XIC(T11_AIRSG2.DN) ,XIC(T12_DLY_TR.DN) ,XIO(T12_DLY_TR.EN) XIC(T12_DLY_TR3.DN) ,XIC(T13_DLY_TR.DN) ,XIO(T13_DLY_TR.EN) XIC(T13_DLY_TR3.DN) ,XIC(T14_DLY_TR.DN) ,XIO(T14_DLY_TR.EN) XIC(T14_DLY_TR3.DN) ,XIC(T15_TRT_ON.DN) ,XIO(T15_TRT_ON.EN) XIC(T15_TRT_OF.DN) ,XIC(T16_TRT_ON.DN) ,XIO(T16_TRT_ON.EN) XIC(T16_TRT_OF.DN) ,XIC(T17_TRT_ON.DN) ,XIO(T17_TRT_ON.EN) XIC(T17_TRT_OF.DN) ,XIC(T21_TRT_ON.DN) ,XIO(T21_TRT_ON.EN) XIC(T21_TRT_OF.DN) ,XIC(T22_TRT_ON.DN) ,XIO(T22_TRT_ON.EN) XIC(T22_TRT_OF.DN) ,XIC(T23_TRT_ON.DN) ,XIO(T23_TRT_ON.EN) XIC(T23_TRT_OF.DN) ,XIC(T24_TRT_ON.DN) ,XIO(T24_TRT_ON.EN) XIC(T24_TRT_OF.DN) ,XIC(T25_TRT_ON.DN) ,XIO(T25_TRT_ON.EN) XIC(T25_TRT_OF.DN) ,XIC(T26_TRT_ON.DN) ,XIO(T26_TRT_ON.EN) XIC(T26_TRT_OF.DN) ,XIC(T27_TRT_ON.DN) ,XIO(T27_TRT_ON.EN) XIC(T27_TRT_OF.DN) ,XIC(T28_TRT_ON.DN) ,XIO(T28_TRT_ON.EN) XIC(T28_TRT_OF.DN) ,XIC(T29_TRT_ON.DN) ,XIO(T29_TRT_ON.EN) XIC(T29_TRT_OF.DN) ,XIC(_709G_TREAT) XIC(_700_TREAT) ][XIC(B9[9].11) ,XIC(B9[9].12) ]XIO(T11_AUTO_A.DN)OTE(O24_007_Bit05);
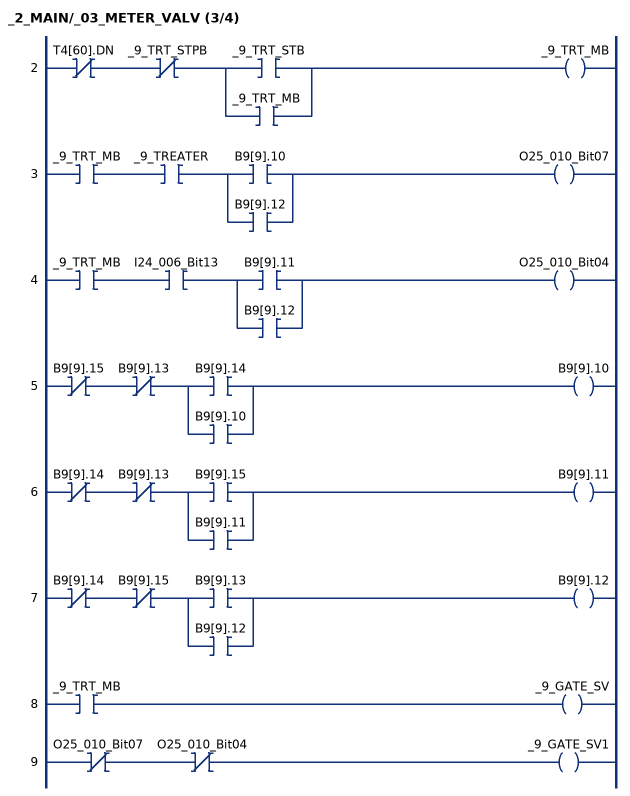
   2: XIO(T4[60].DN)XIO(_9_TRT_STPB)[XIC(_9_TRT_STB) ,XIC(_9_TRT_MB) ]OTE(_9_TRT_MB);
   3: XIC(_9_TRT_MB)XIC(_9_TREATER)[XIC(B9[9].10) ,XIC(B9[9].12) ]OTE(O25_010_Bit07);
   4: XIC(_9_TRT_MB)XIC(I24_006_Bit13)[XIC(B9[9].11) ,XIC(B9[9].12) ]OTE(O25_010_Bit04);
   5: XIO(B9[9].15)XIO(B9[9].13)[XIC(B9[9].14) ,XIC(B9[9].10) ]OTE(B9[9].10);
   6: XIO(B9[9].14)XIO(B9[9].13)[XIC(B9[9].15) ,XIC(B9[9].11) ]OTE(B9[9].11);
   7: XIO(B9[9].14)XIO(B9[9].15)[XIC(B9[9].13) ,XIC(B9[9].12) ]OTE(B9[9].12);
   8: XIC(_9_TRT_MB)OTE(_9_GATE_SV);
   9: XIO(O25_010_Bit07)XIO(O25_010_Bit04)OTE(_9_GATE_SV1);
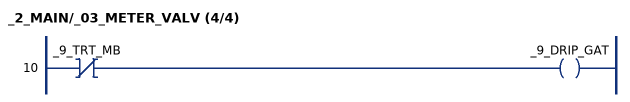
   10: XIO(_9_TRT_MB)OTE(_9_DRIP_GAT);
END_ROUTINE

ROUTINE _04_TREAT_DELY   (* ladder *)
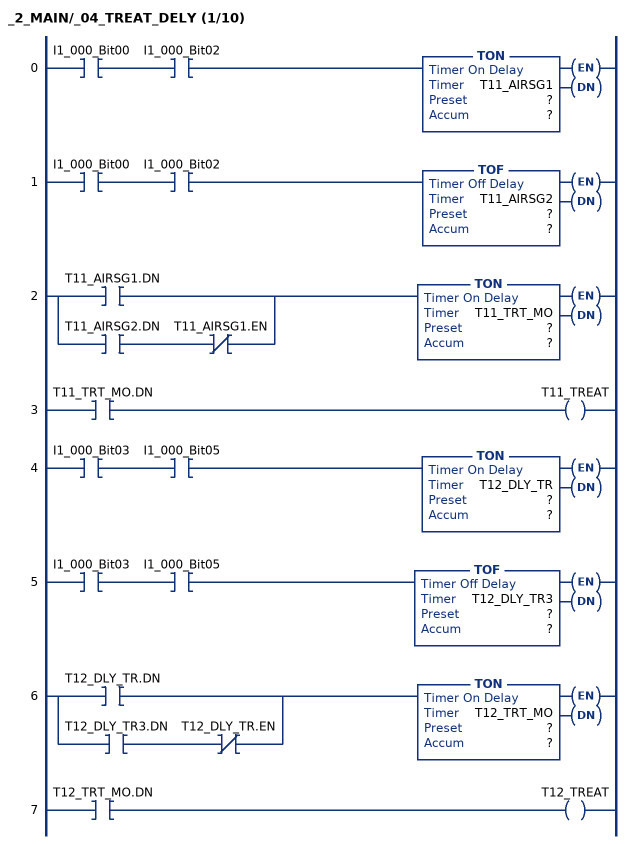
   0: XIC(I1_000_Bit00)XIC(I1_000_Bit02)TON(T11_AIRSG1,?,?);
   1: XIC(I1_000_Bit00)XIC(I1_000_Bit02)TOF(T11_AIRSG2,?,?);
   2: [XIC(T11_AIRSG1.DN) ,XIC(T11_AIRSG2.DN) XIO(T11_AIRSG1.EN) ]TON(T11_TRT_MO,?,?);
   3: XIC(T11_TRT_MO.DN)OTE(T11_TREAT);
   4: XIC(I1_000_Bit03)XIC(I1_000_Bit05)TON(T12_DLY_TR,?,?);
   5: XIC(I1_000_Bit03)XIC(I1_000_Bit05)TOF(T12_DLY_TR3,?,?);
   6: [XIC(T12_DLY_TR.DN) ,XIC(T12_DLY_TR3.DN) XIO(T12_DLY_TR.EN) ]TON(T12_TRT_MO,?,?);
   7: XIC(T12_TRT_MO.DN)OTE(T12_TREAT);
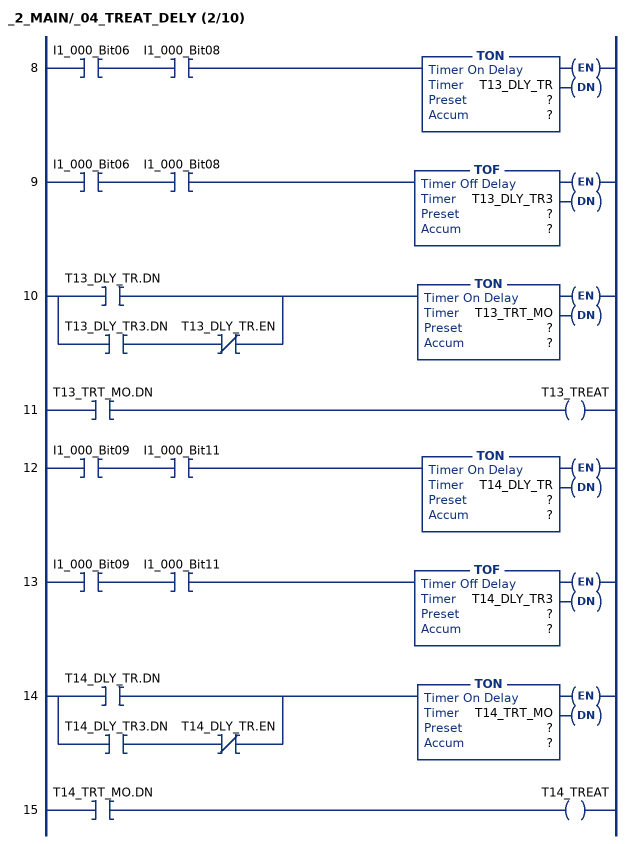
   8: XIC(I1_000_Bit06)XIC(I1_000_Bit08)TON(T13_DLY_TR,?,?);
   9: XIC(I1_000_Bit06)XIC(I1_000_Bit08)TOF(T13_DLY_TR3,?,?);
   10: [XIC(T13_DLY_TR.DN) ,XIC(T13_DLY_TR3.DN) XIO(T13_DLY_TR.EN) ]TON(T13_TRT_MO,?,?);
   11: XIC(T13_TRT_MO.DN)OTE(T13_TREAT);
   12: XIC(I1_000_Bit09)XIC(I1_000_Bit11)TON(T14_DLY_TR,?,?);
   13: XIC(I1_000_Bit09)XIC(I1_000_Bit11)TOF(T14_DLY_TR3,?,?);
   14: [XIC(T14_DLY_TR.DN) ,XIC(T14_DLY_TR3.DN) XIO(T14_DLY_TR.EN) ]TON(T14_TRT_MO,?,?);
   15: XIC(T14_TRT_MO.DN)OTE(T14_TREAT);
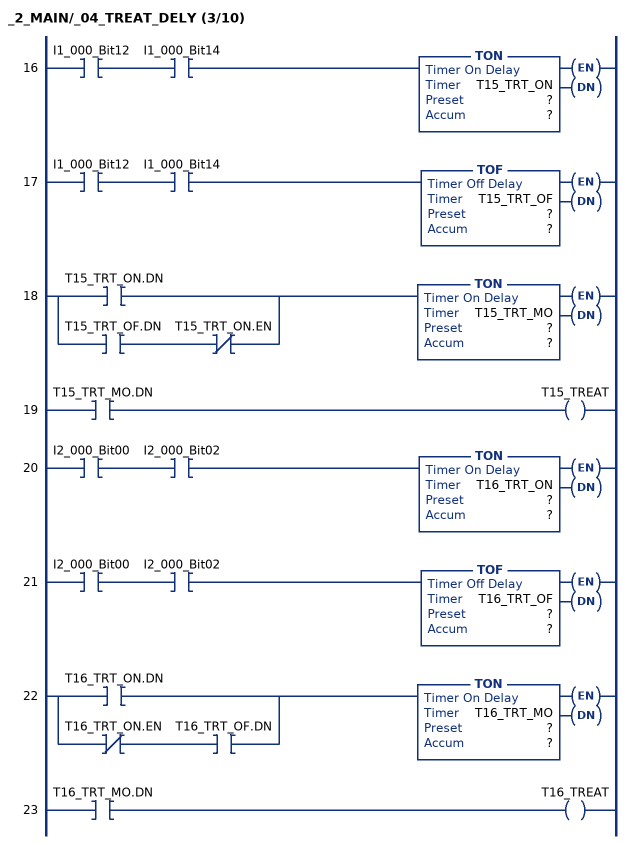
   16: XIC(I1_000_Bit12)XIC(I1_000_Bit14)TON(T15_TRT_ON,?,?);
   17: XIC(I1_000_Bit12)XIC(I1_000_Bit14)TOF(T15_TRT_OF,?,?);
   18: [XIC(T15_TRT_ON.DN) ,XIC(T15_TRT_OF.DN) XIO(T15_TRT_ON.EN) ]TON(T15_TRT_MO,?,?);
   19: XIC(T15_TRT_MO.DN)OTE(T15_TREAT);
   20: XIC(I2_000_Bit00)XIC(I2_000_Bit02)TON(T16_TRT_ON,?,?);
   21: XIC(I2_000_Bit00)XIC(I2_000_Bit02)TOF(T16_TRT_OF,?,?);
   22: [XIC(T16_TRT_ON.DN) ,XIO(T16_TRT_ON.EN) XIC(T16_TRT_OF.DN) ]TON(T16_TRT_MO,?,?);
   23: XIC(T16_TRT_MO.DN)OTE(T16_TREAT);
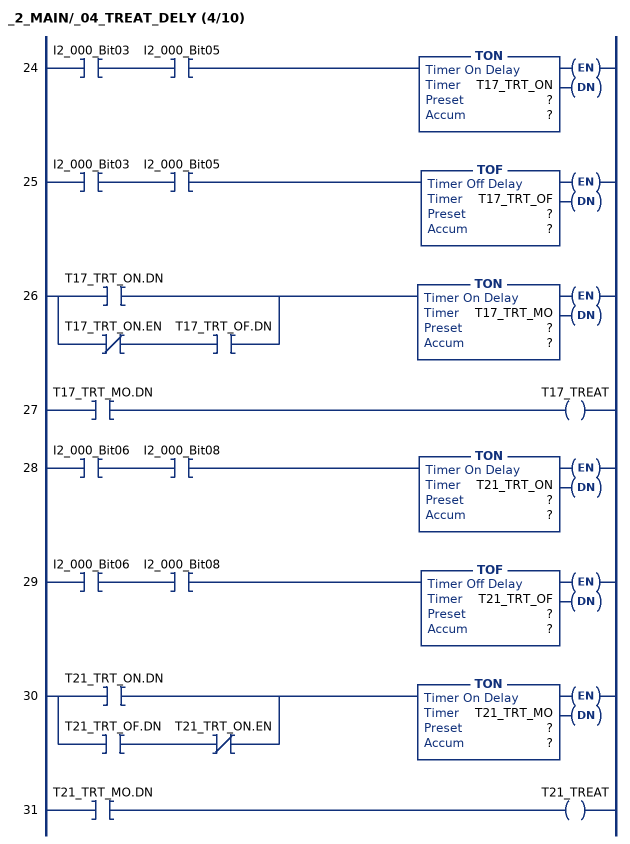
   24: XIC(I2_000_Bit03)XIC(I2_000_Bit05)TON(T17_TRT_ON,?,?);
   25: XIC(I2_000_Bit03)XIC(I2_000_Bit05)TOF(T17_TRT_OF,?,?);
   26: [XIC(T17_TRT_ON.DN) ,XIO(T17_TRT_ON.EN) XIC(T17_TRT_OF.DN) ]TON(T17_TRT_MO,?,?);
   27: XIC(T17_TRT_MO.DN)OTE(T17_TREAT);
   28: XIC(I2_000_Bit06)XIC(I2_000_Bit08)TON(T21_TRT_ON,?,?);
   29: XIC(I2_000_Bit06)XIC(I2_000_Bit08)TOF(T21_TRT_OF,?,?);
   30: [XIC(T21_TRT_ON.DN) ,XIC(T21_TRT_OF.DN) XIO(T21_TRT_ON.EN) ]TON(T21_TRT_MO,?,?);
   31: XIC(T21_TRT_MO.DN)OTE(T21_TREAT);
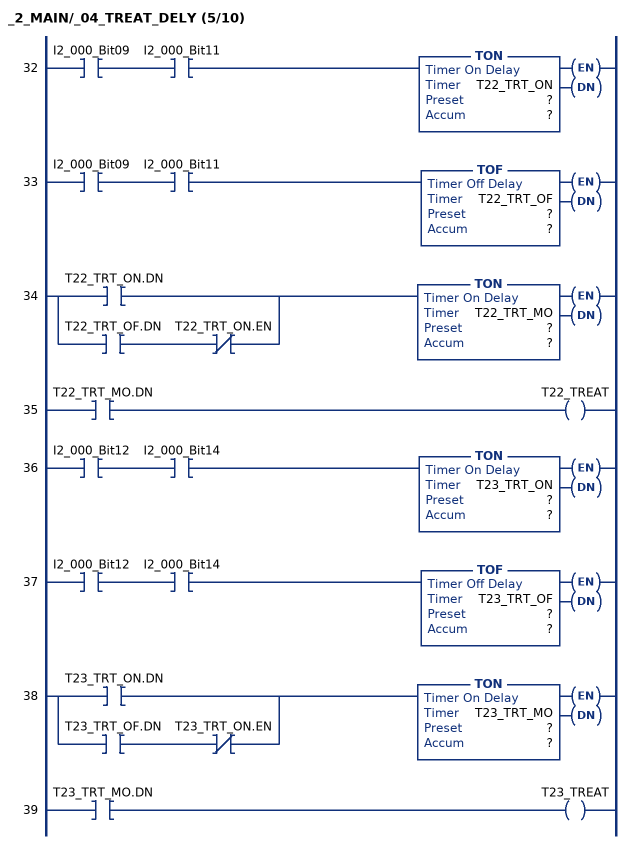
   32: XIC(I2_000_Bit09)XIC(I2_000_Bit11)TON(T22_TRT_ON,?,?);
   33: XIC(I2_000_Bit09)XIC(I2_000_Bit11)TOF(T22_TRT_OF,?,?);
   34: [XIC(T22_TRT_ON.DN) ,XIC(T22_TRT_OF.DN) XIO(T22_TRT_ON.EN) ]TON(T22_TRT_MO,?,?);
   35: XIC(T22_TRT_MO.DN)OTE(T22_TREAT);
   36: XIC(I2_000_Bit12)XIC(I2_000_Bit14)TON(T23_TRT_ON,?,?);
   37: XIC(I2_000_Bit12)XIC(I2_000_Bit14)TOF(T23_TRT_OF,?,?);
   38: [XIC(T23_TRT_ON.DN) ,XIC(T23_TRT_OF.DN) XIO(T23_TRT_ON.EN) ]TON(T23_TRT_MO,?,?);
   39: XIC(T23_TRT_MO.DN)OTE(T23_TREAT);
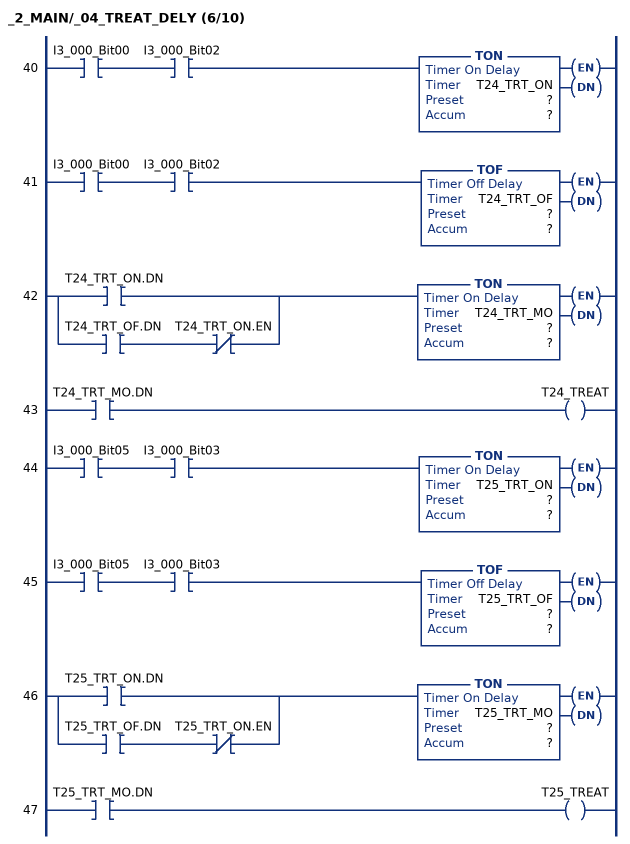
   40: XIC(I3_000_Bit00)XIC(I3_000_Bit02)TON(T24_TRT_ON,?,?);
   41: XIC(I3_000_Bit00)XIC(I3_000_Bit02)TOF(T24_TRT_OF,?,?);
   42: [XIC(T24_TRT_ON.DN) ,XIC(T24_TRT_OF.DN) XIO(T24_TRT_ON.EN) ]TON(T24_TRT_MO,?,?);
   43: XIC(T24_TRT_MO.DN)OTE(T24_TREAT);
   44: XIC(I3_000_Bit05)XIC(I3_000_Bit03)TON(T25_TRT_ON,?,?);
   45: XIC(I3_000_Bit05)XIC(I3_000_Bit03)TOF(T25_TRT_OF,?,?);
   46: [XIC(T25_TRT_ON.DN) ,XIC(T25_TRT_OF.DN) XIO(T25_TRT_ON.EN) ]TON(T25_TRT_MO,?,?);
   47: XIC(T25_TRT_MO.DN)OTE(T25_TREAT);
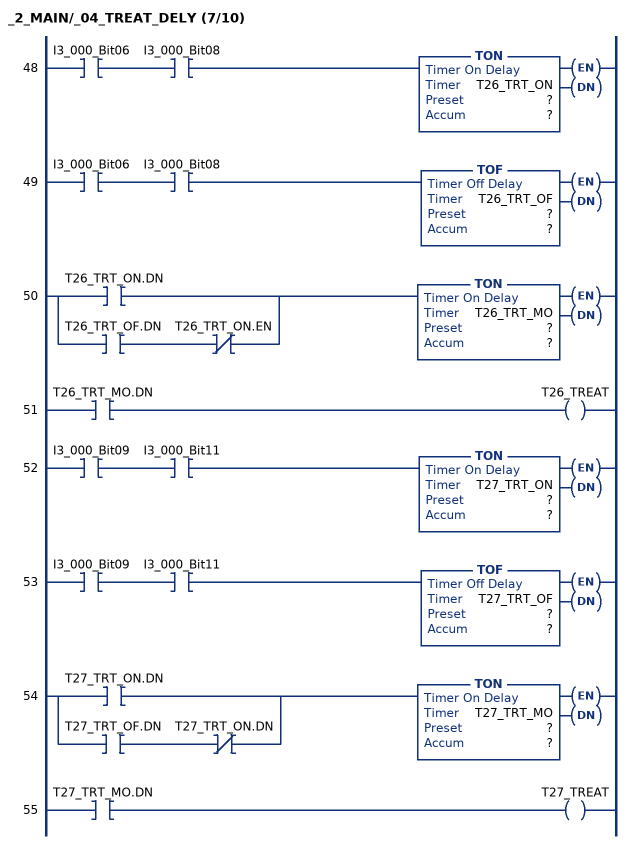
   48: XIC(I3_000_Bit06)XIC(I3_000_Bit08)TON(T26_TRT_ON,?,?);
   49: XIC(I3_000_Bit06)XIC(I3_000_Bit08)TOF(T26_TRT_OF,?,?);
   50: [XIC(T26_TRT_ON.DN) ,XIC(T26_TRT_OF.DN) XIO(T26_TRT_ON.EN) ]TON(T26_TRT_MO,?,?);
   51: XIC(T26_TRT_MO.DN)OTE(T26_TREAT);
   52: XIC(I3_000_Bit09)XIC(I3_000_Bit11)TON(T27_TRT_ON,?,?);
   53: XIC(I3_000_Bit09)XIC(I3_000_Bit11)TOF(T27_TRT_OF,?,?);
   54: [XIC(T27_TRT_ON.DN) ,XIC(T27_TRT_OF.DN) XIO(T27_TRT_ON.DN) ]TON(T27_TRT_MO,?,?);
   55: XIC(T27_TRT_MO.DN)OTE(T27_TREAT);
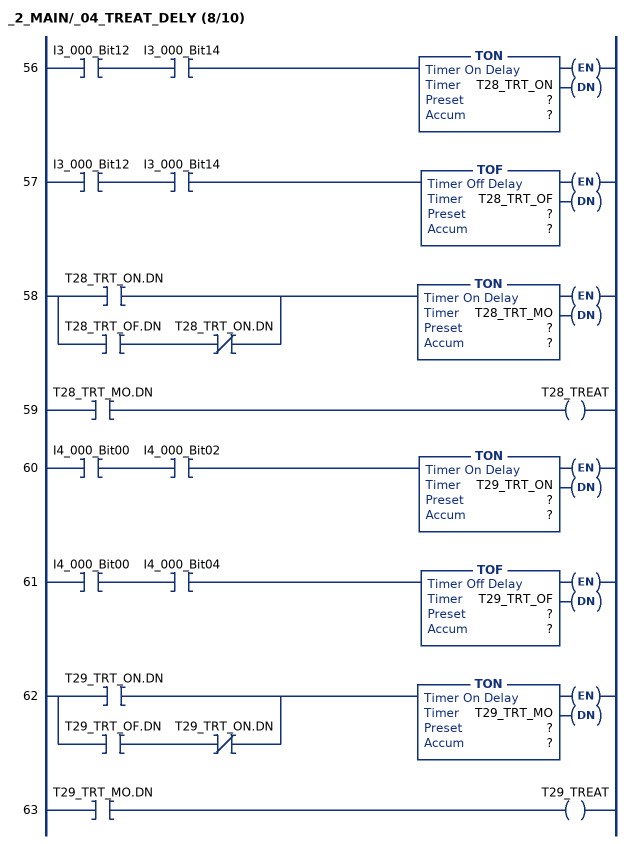
   56: XIC(I3_000_Bit12)XIC(I3_000_Bit14)TON(T28_TRT_ON,?,?);
   57: XIC(I3_000_Bit12)XIC(I3_000_Bit14)TOF(T28_TRT_OF,?,?);
   58: [XIC(T28_TRT_ON.DN) ,XIC(T28_TRT_OF.DN) XIO(T28_TRT_ON.DN) ]TON(T28_TRT_MO,?,?);
   59: XIC(T28_TRT_MO.DN)OTE(T28_TREAT);
   60: XIC(I4_000_Bit00)XIC(I4_000_Bit02)TON(T29_TRT_ON,?,?);
   61: XIC(I4_000_Bit00)XIC(I4_000_Bit04)TOF(T29_TRT_OF,?,?);
   62: [XIC(T29_TRT_ON.DN) ,XIC(T29_TRT_OF.DN) XIO(T29_TRT_ON.DN) ]TON(T29_TRT_MO,?,?);
   63: XIC(T29_TRT_MO.DN)OTE(T29_TREAT);
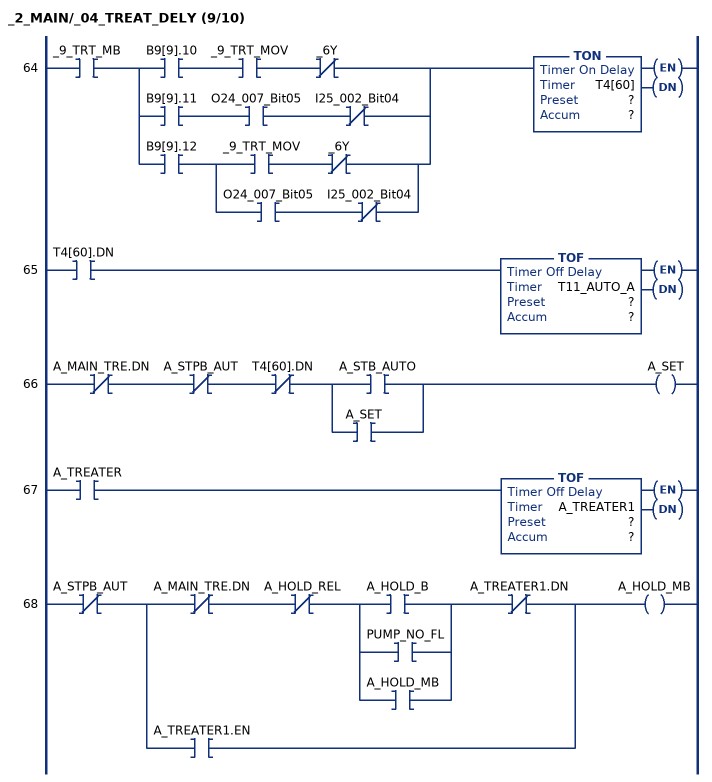
   64: XIC(_9_TRT_MB)[XIC(B9[9].10) XIC(_9_TRT_MOV) XIO(_6Y) ,XIC(B9[9].11) XIC(O24_007_Bit05) XIO(I25_002_Bit04) ,XIC(B9[9].12) [XIC(_9_TRT_MOV) XIO(_6Y) ,XIC(O24_007_Bit05) XIO(I25_002_Bit04) ] ]TON(T4[60],?,?);
   65: XIC(T4[60].DN)TOF(T11_AUTO_A,?,?);
   66: XIO(A_MAIN_TRE.DN)XIO(A_STPB_AUT)XIO(T4[60].DN)[XIC(A_STB_AUTO) ,XIC(A_SET) ]OTE(A_SET);
   67: XIC(A_TREATER)TOF(A_TREATER1,?,?);
   68: XIO(A_STPB_AUT)[XIO(A_MAIN_TRE.DN) XIO(A_HOLD_REL) [XIC(A_HOLD_B) ,XIC(PUMP_NO_FL) ,XIC(A_HOLD_MB) ] XIO(A_TREATER1.DN) ,XIC(A_TREATER1.EN) ]OTE(A_HOLD_MB);
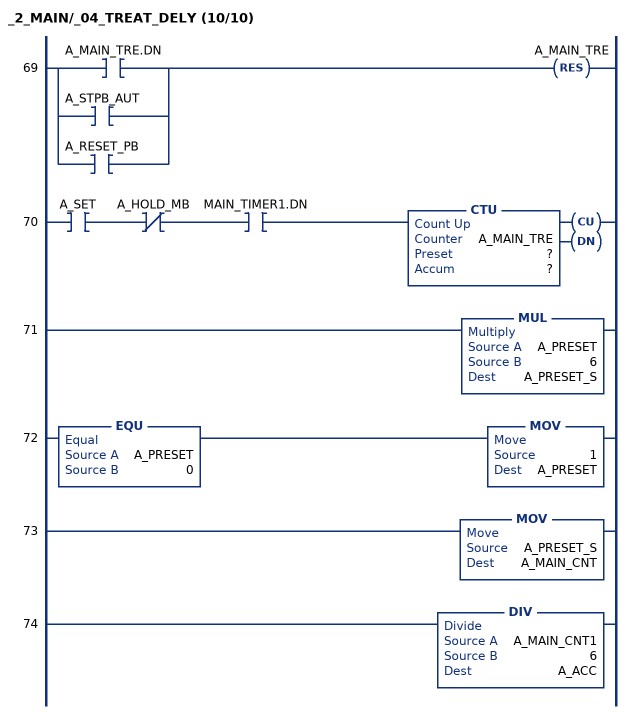
   69: [XIC(A_MAIN_TRE.DN) ,XIC(A_STPB_AUT) ,XIC(A_RESET_PB) ]RES(A_MAIN_TRE);
   70: XIC(A_SET)XIO(A_HOLD_MB)XIC(MAIN_TIMER1.DN)CTU(A_MAIN_TRE,?,?);
   71: MUL(A_PRESET,6,A_PRESET_S);
   72: EQU(A_PRESET,0)MOV(1,A_PRESET);
   73: MOV(A_PRESET_S,A_MAIN_CNT);
   74: DIV(A_MAIN_CNT1,6,A_ACC);
END_ROUTINE

ROUTINE _05_5_PMPS_ATO   (* ladder *)
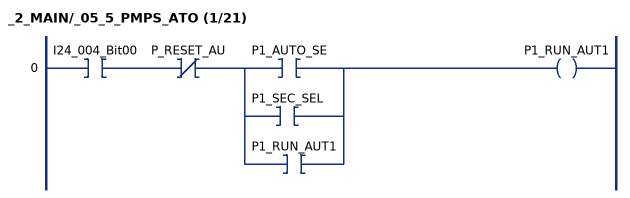
   0: XIC(I24_004_Bit00)XIO(P_RESET_AU)[XIC(P1_AUTO_SE) ,XIC(P1_SEC_SEL) ,XIC(P1_RUN_AUT1) ]OTE(P1_RUN_AUT1);
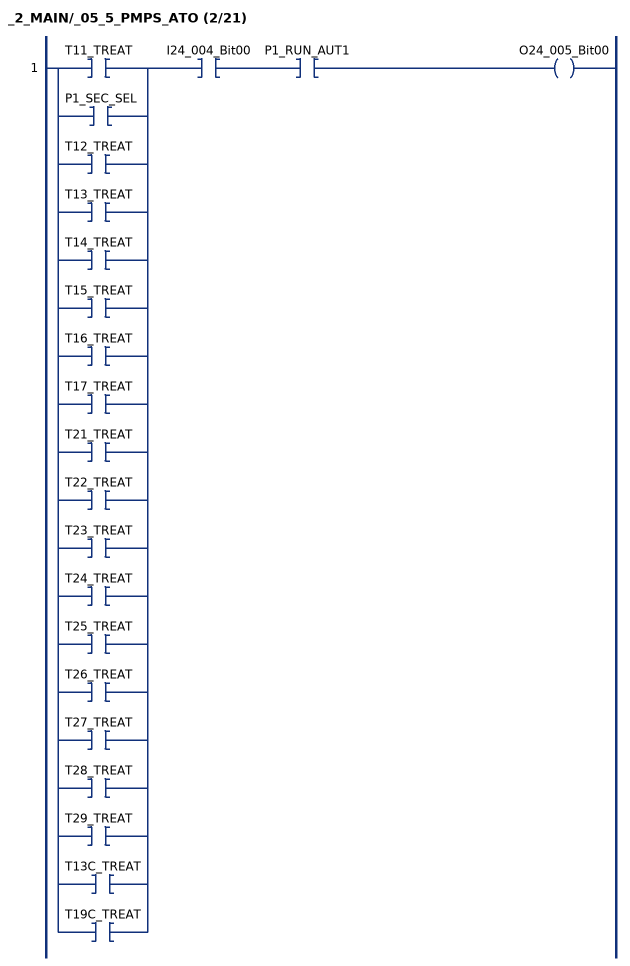
   1: [XIC(T11_TREAT) ,XIC(P1_SEC_SEL) ,XIC(T12_TREAT) ,XIC(T13_TREAT) ,XIC(T14_TREAT) ,XIC(T15_TREAT) ,XIC(T16_TREAT) ,XIC(T17_TREAT) ,XIC(T21_TREAT) ,XIC(T22_TREAT) ,XIC(T23_TREAT) ,XIC(T24_TREAT) ,XIC(T25_TREAT) ,XIC(T26_TREAT) ,XIC(T27_TREAT) ,XIC(T28_TREAT) ,XIC(T29_TREAT) ,XIC(T13C_TREAT) ,XIC(T19C_TREAT) ]XIC(I24_004_Bit00)XIC(P1_RUN_AUT1)OTE(O24_005_Bit00);
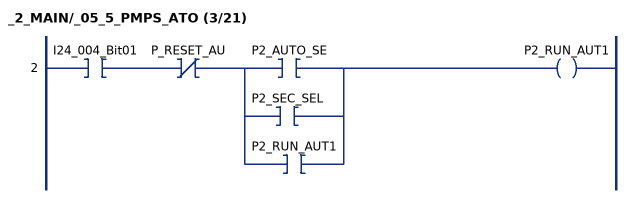
   2: XIC(I24_004_Bit01)XIO(P_RESET_AU)[XIC(P2_AUTO_SE) ,XIC(P2_SEC_SEL) ,XIC(P2_RUN_AUT1) ]OTE(P2_RUN_AUT1);
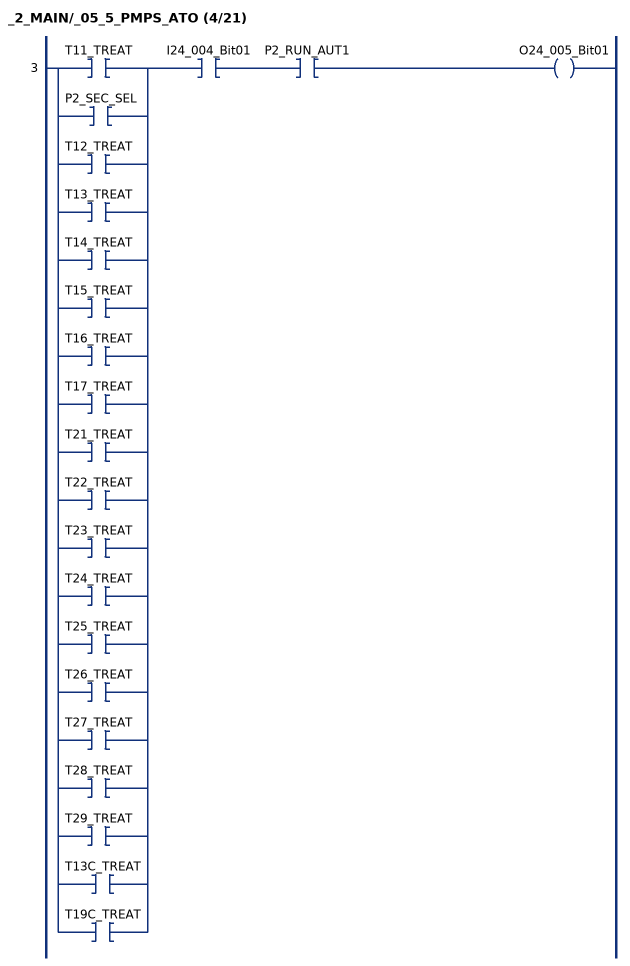
   3: [XIC(T11_TREAT) ,XIC(P2_SEC_SEL) ,XIC(T12_TREAT) ,XIC(T13_TREAT) ,XIC(T14_TREAT) ,XIC(T15_TREAT) ,XIC(T16_TREAT) ,XIC(T17_TREAT) ,XIC(T21_TREAT) ,XIC(T22_TREAT) ,XIC(T23_TREAT) ,XIC(T24_TREAT) ,XIC(T25_TREAT) ,XIC(T26_TREAT) ,XIC(T27_TREAT) ,XIC(T28_TREAT) ,XIC(T29_TREAT) ,XIC(T13C_TREAT) ,XIC(T19C_TREAT) ]XIC(I24_004_Bit01)XIC(P2_RUN_AUT1)OTE(O24_005_Bit01);
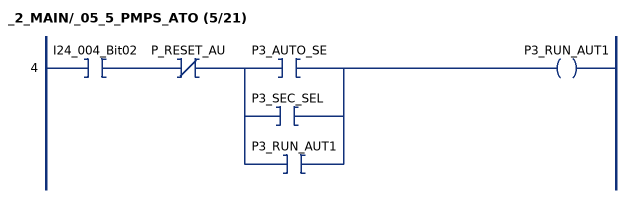
   4: XIC(I24_004_Bit02)XIO(P_RESET_AU)[XIC(P3_AUTO_SE) ,XIC(P3_SEC_SEL) ,XIC(P3_RUN_AUT1) ]OTE(P3_RUN_AUT1);
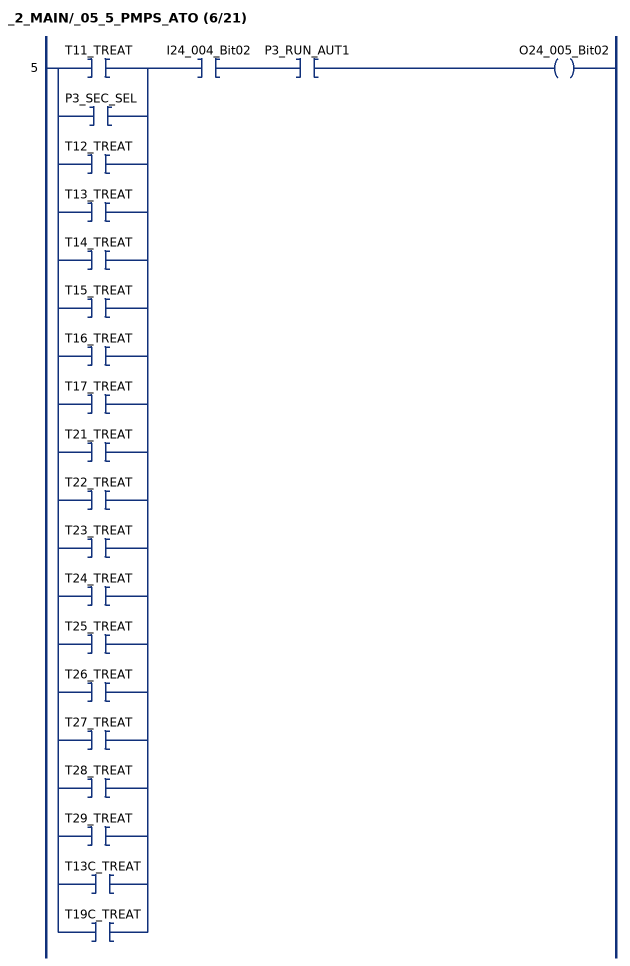
   5: [XIC(T11_TREAT) ,XIC(P3_SEC_SEL) ,XIC(T12_TREAT) ,XIC(T13_TREAT) ,XIC(T14_TREAT) ,XIC(T15_TREAT) ,XIC(T16_TREAT) ,XIC(T17_TREAT) ,XIC(T21_TREAT) ,XIC(T22_TREAT) ,XIC(T23_TREAT) ,XIC(T24_TREAT) ,XIC(T25_TREAT) ,XIC(T26_TREAT) ,XIC(T27_TREAT) ,XIC(T28_TREAT) ,XIC(T29_TREAT) ,XIC(T13C_TREAT) ,XIC(T19C_TREAT) ]XIC(I24_004_Bit02)XIC(P3_RUN_AUT1)OTE(O24_005_Bit02);
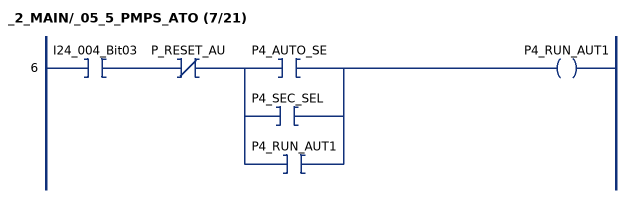
   6: XIC(I24_004_Bit03)XIO(P_RESET_AU)[XIC(P4_AUTO_SE) ,XIC(P4_SEC_SEL) ,XIC(P4_RUN_AUT1) ]OTE(P4_RUN_AUT1);
